PatternFound := FALSE;
IF ExpectedLength = USINT_TO_DINT(Length) THEN
    LastCandidateOffset := 0;
    FOR CandidateOffset := 0 TO LastCandidateOffset DO
        PatternMatches := TRUE;
        FOR CharacterIndex := 0 TO ExpectedLength - 1 DO
            InIndex := LINT_TO_DINT(DINT_TO_LINT(StartIndex) + CandidateOffset
                + DINT_TO_LINT(CharacterIndex));
            IF IN[InIndex] <> Expected[CharacterIndex] THEN
                PatternMatches := FALSE;
                EXIT;
            END_IF;
        END_FOR;
        IF PatternMatches THEN
            PatternFound := TRUE;
            EXIT;
        END_IF;
    END_FOR;
END_IF;

IF NOT PatternFound THEN
    ExpectedText := CreateAssertionTextValue_WString(Value := Expected);
    Message := CONCAT('Assertion failed: selected array does not equal Expected = ',
        ExpectedText);
    Message := CONCAT(Message, ', Range = [');
    Message := CONCAT(Message, DINT_TO_STRING(StartIndex));
    Message := CONCAT(Message, '..');
    Message := CONCAT(Message, LINT_TO_STRING(EndIndex));
    Message := CONCAT(Message, '], ExpectedLength = ');
    Message := CONCAT(Message, DINT_TO_STRING(ExpectedLength));
    Message := CONCAT(Message, '.');
    Fail(Message := Message);
    RETURN;
END_IF;

Pass();
{warning restore C0371}
END_METHOD

END_FUNCTION_BLOCK

// ---- Framework/Assertions/POU/Utilities/IsAssertionWStringLengthValid.TcPOU
{region 'Documentation'}
(*!
<summary>Checks for a terminator within the configured content capacity, including empty text. Reads at most capacity + 1 code units and stops at the first terminator.</summary>
*)
{endregion}
FUNCTION INTERNAL IsAssertionWStringLengthValid : BOOL //! TRUE when a terminator occurs within the configured capacity, including empty text.
VAR_IN_OUT CONSTANT
    Value : WSTRING(Param_Assertions.AssertionWStringLength); //! Read-only text to check for termination within its configured capacity.
END_VAR
VAR
    CharacterIndex : DINT;
END_VAR
VAR CONSTANT
    Terminator : WORD := 0;
END_VAR

IsAssertionWStringLengthValid := FALSE;
FOR CharacterIndex := 0 TO UINT_TO_DINT(Param_Assertions.AssertionWStringLength) DO
    IF Value[CharacterIndex] = Terminator THEN
        IsAssertionWStringLengthValid := TRUE;
        RETURN;
    END_IF;
END_FOR;

END_FUNCTION

// ---- Framework/Assertions/POU/Arrays/Word/AssertArrayContainsWString_Word.TcPOU
{region 'Documentation'}
(*!
<summary>Search the selected array for the contiguous WSTRING code units.</summary>
<description>

StartIndex is an absolute declared IN index, not an offset. Length selects 1..255
elements; the complete selected range must fit IN. Invalid references or ranges report
Error.

Keep supplied arrays stable for the call. Input data is read, not copied or retained as a
snapshot.

Expected must be nonempty and fit its configured text capacity (otherwise Error). A valid
text longer than the selected array region reports Failed. The array is not zero-terminated or
trimmed; matching is exact and case-sensitive.

</description>
*)
{endregion}
FUNCTION_BLOCK AssertArrayContainsWString_Word EXTENDS AssertionBase
VAR_INPUT
    StartIndex : DINT; //! First selected index in IN; uses the array's declared index range, not a zero-based offset.
    Length : USINT; //! Number of selected array elements, from 1 through 255.
END_VAR
VAR_IN_OUT CONSTANT
    IN : ARRAY[*] OF WORD; //! Read-only actual data; the selected range must remain stable during the call.
    Expected : WSTRING(Param_Assertions.AssertionWStringLength); //! Nonempty expected text, terminated within the configured capacity; keep stable during the call.
END_VAR

SUPER^();

{region 'Documentation'}
(*!
<summary>Validate references and ranges before exact code-unit comparison.</summary>
*)
{endregion}
METHOD PROTECTED Assert
VAR
    InLowerIndex : DINT;
    InUpperIndex : DINT;
    EndIndex : LINT;
    ExpectedLength : DINT;
    CharacterIndex : DINT;
    InIndex : DINT;
    CandidateOffset : LINT;
    LastCandidateOffset : LINT;
    PatternMatches : BOOL;
    PatternFound : BOOL;
    ExpectedText : STRING(GVL_Constants.AssertionValueLength);
    Message : STRING(GVL_Constants.MessageLength);
END_VAR
VAR CONSTANT
    Terminator : WORD := 0;
END_VAR
IF NOT EvaluationActive THEN
    RETURN;
END_IF;

IF Result = E_Result.Error THEN
    RETURN;
END_IF;

// C0371: FB inputs are checked before any reference access.
{warning disable C0371}
IF NOT __ISVALIDREF(IN) THEN
    Error(Message := 'Assertion error: IN reference is invalid.');
    RETURN;
END_IF;

IF NOT __ISVALIDREF(Expected) THEN
    Error(Message := 'Assertion error: Expected reference is invalid.');
    RETURN;
END_IF;

IF NOT IsAssertionWStringLengthValid(Value := Expected) THEN
    Error(Message := 'Assertion error: Expected exceeds configured WSTRING length.');
    RETURN;
END_IF;

IF Expected[0] = Terminator THEN
    Error(Message := 'Assertion error: Expected must not be empty.');
    RETURN;
END_IF;

ExpectedLength := 0;
FOR CharacterIndex := 0 TO UINT_TO_DINT(Param_Assertions.AssertionWStringLength) DO
    IF Expected[CharacterIndex] = Terminator THEN
        ExpectedLength := CharacterIndex;
        EXIT;
    END_IF;
END_FOR;

InLowerIndex := LOWER_BOUND(IN, 1);
InUpperIndex := UPPER_BOUND(IN, 1);
EndIndex := DINT_TO_LINT(StartIndex) + USINT_TO_LINT(Length) - 1;
IF (Length = 0)
    OR (StartIndex < InLowerIndex) OR (StartIndex > InUpperIndex)
    OR (EndIndex > DINT_TO_LINT(InUpperIndex)) THEN
    Message := CONCAT('Assertion error: array range is invalid. StartIndex = ',
        DINT_TO_STRING(StartIndex));
    Message := CONCAT(Message, ', Length = ');
    Message := CONCAT(Message, USINT_TO_STRING(Length));
    Error(Message := Message);
    RETURN;
END_IF;

IF Result = E_Result.Failed THEN
    RETURN;
END_IF;

PatternFound := FALSE;
IF ExpectedLength <= USINT_TO_DINT(Length) THEN
    LastCandidateOffset := USINT_TO_LINT(Length) - DINT_TO_LINT(ExpectedLength);
    FOR CandidateOffset := 0 TO LastCandidateOffset DO
        PatternMatches := TRUE;
        FOR CharacterIndex := 0 TO ExpectedLength - 1 DO
            InIndex := LINT_TO_DINT(DINT_TO_LINT(StartIndex) + CandidateOffset
                + DINT_TO_LINT(CharacterIndex));
            IF IN[InIndex] <> Expected[CharacterIndex] THEN
                PatternMatches := FALSE;
                EXIT;
            END_IF;
        END_FOR;
        IF PatternMatches THEN
            PatternFound := TRUE;
            EXIT;
        END_IF;
    END_FOR;
END_IF;

IF NOT PatternFound THEN
    ExpectedText := CreateAssertionTextValue_WString(Value := Expected);
    Message := CONCAT('Assertion failed: selected array does not contain Expected = ',
        ExpectedText);
    Message := CONCAT(Message, ', Range = [');
    Message := CONCAT(Message, DINT_TO_STRING(StartIndex));
    Message := CONCAT(Message, '..');
    Message := CONCAT(Message, LINT_TO_STRING(EndIndex));
    Message := CONCAT(Message, '], ExpectedLength = ');
    Message := CONCAT(Message, DINT_TO_STRING(ExpectedLength));
    Message := CONCAT(Message, '.');
    Fail(Message := Message);
    RETURN;
END_IF;

Pass();
{warning restore C0371}
END_METHOD

END_FUNCTION_BLOCK

// ---- Framework/Assertions/POU/Arrays/Word/AssertArrayStartsWithWString_Word.TcPOU
{region 'Documentation'}
(*!
<summary>Check that the selected array starts with the WSTRING code units.</summary>
<description>

StartIndex is an absolute declared IN index, not an offset. Length selects 1..255
elements; the complete selected range must fit IN. Invalid references or ranges report
Error.

Keep supplied arrays stable for the call. Input data is read, not copied or retained as a
snapshot.

Expected must be nonempty and fit its configured text capacity (otherwise Error). A valid
text longer than the selected array region reports Failed. The array is not zero-terminated or
trimmed; matching is exact and case-sensitive.

</description>
*)
{endregion}
FUNCTION_BLOCK AssertArrayStartsWithWString_Word EXTENDS AssertionBase
VAR_INPUT
    StartIndex : DINT; //! First selected index in IN; uses the array's declared index range, not a zero-based offset.
    Length : USINT; //! Number of selected array elements, from 1 through 255.
END_VAR
VAR_IN_OUT CONSTANT
    IN : ARRAY[*] OF WORD; //! Read-only actual data; the selected range must remain stable during the call.
    Expected : WSTRING(Param_Assertions.AssertionWStringLength); //! Nonempty expected text, terminated within the configured capacity; keep stable during the call.
END_VAR

SUPER^();

{region 'Documentation'}
(*!
<summary>Validate references and ranges before exact code-unit comparison.</summary>
*)
{endregion}
METHOD PROTECTED Assert
VAR
    InLowerIndex : DINT;
    InUpperIndex : DINT;
    EndIndex : LINT;
    ExpectedLength : DINT;
    CharacterIndex : DINT;
    InIndex : DINT;
    CandidateOffset : LINT;
    LastCandidateOffset : LINT;
    PatternMatches : BOOL;
    PatternFound : BOOL;
    ExpectedText : STRING(GVL_Constants.AssertionValueLength);
    Message : STRING(GVL_Constants.MessageLength);
END_VAR
VAR CONSTANT
    Terminator : WORD := 0;
END_VAR
IF NOT EvaluationActive THEN
    RETURN;
END_IF;

IF Result = E_Result.Error THEN
    RETURN;
END_IF;

// C0371: FB inputs are checked before any reference access.
{warning disable C0371}
IF NOT __ISVALIDREF(IN) THEN
    Error(Message := 'Assertion error: IN reference is invalid.');
    RETURN;
END_IF;

IF NOT __ISVALIDREF(Expected) THEN
    Error(Message := 'Assertion error: Expected reference is invalid.');
    RETURN;
END_IF;

IF NOT IsAssertionWStringLengthValid(Value := Expected) THEN
    Error(Message := 'Assertion error: Expected exceeds configured WSTRING length.');
    RETURN;
END_IF;

IF Expected[0] = Terminator THEN
    Error(Message := 'Assertion error: Expected must not be empty.');
    RETURN;
END_IF;

ExpectedLength := 0;
FOR CharacterIndex := 0 TO UINT_TO_DINT(Param_Assertions.AssertionWStringLength) DO
    IF Expected[CharacterIndex] = Terminator THEN
        ExpectedLength := CharacterIndex;
        EXIT;
    END_IF;
END_FOR;

InLowerIndex := LOWER_BOUND(IN, 1);
InUpperIndex := UPPER_BOUND(IN, 1);
EndIndex := DINT_TO_LINT(StartIndex) + USINT_TO_LINT(Length) - 1;
IF (Length = 0)
    OR (StartIndex < InLowerIndex) OR (StartIndex > InUpperIndex)
    OR (EndIndex > DINT_TO_LINT(InUpperIndex)) THEN
    Message := CONCAT('Assertion error: array range is invalid. StartIndex = ',
        DINT_TO_STRING(StartIndex));
    Message := CONCAT(Message, ', Length = ');
    Message := CONCAT(Message, USINT_TO_STRING(Length));
    Error(Message := Message);
    RETURN;
END_IF;

IF Result = E_Result.Failed THEN
    RETURN;
END_IF;

PatternFound := FALSE;
IF ExpectedLength <= USINT_TO_DINT(Length) THEN
    LastCandidateOffset := 0;
    FOR CandidateOffset := 0 TO LastCandidateOffset DO
        PatternMatches := TRUE;
        FOR CharacterIndex := 0 TO ExpectedLength - 1 DO
            InIndex := LINT_TO_DINT(DINT_TO_LINT(StartIndex) + CandidateOffset
                + DINT_TO_LINT(CharacterIndex));
            IF IN[InIndex] <> Expected[CharacterIndex] THEN
                PatternMatches := FALSE;
                EXIT;
            END_IF;
        END_FOR;
        IF PatternMatches THEN
            PatternFound := TRUE;
            EXIT;
        END_IF;
    END_FOR;
END_IF;

IF NOT PatternFound THEN
    ExpectedText := CreateAssertionTextValue_WString(Value := Expected);
    Message := CONCAT('Assertion failed: selected array does not start with Expected = ',
        ExpectedText);
    Message := CONCAT(Message, ', Range = [');
    Message := CONCAT(Message, DINT_TO_STRING(StartIndex));
    Message := CONCAT(Message, '..');
    Message := CONCAT(Message, LINT_TO_STRING(EndIndex));
    Message := CONCAT(Message, '], ExpectedLength = ');
    Message := CONCAT(Message, DINT_TO_STRING(ExpectedLength));
    Message := CONCAT(Message, '.');
    Fail(Message := Message);
    RETURN;
END_IF;

Pass();
{warning restore C0371}
END_METHOD

END_FUNCTION_BLOCK

// ---- Framework/Assertions/POU/Arrays/Word/AssertArrayEndsWithWString_Word.TcPOU
{region 'Documentation'}
(*!
<summary>Check that the selected array ends with the WSTRING code units.</summary>
<description>

StartIndex is an absolute declared IN index, not an offset. Length selects 1..255
elements; the complete selected range must fit IN. Invalid references or ranges report
Error.

Keep supplied arrays stable for the call. Input data is read, not copied or retained as a
snapshot.

Expected must be nonempty and fit its configured text capacity (otherwise Error). A valid
text longer than the selected array region reports Failed. The array is not zero-terminated or
trimmed; matching is exact and case-sensitive.

</description>
*)
{endregion}
FUNCTION_BLOCK AssertArrayEndsWithWString_Word EXTENDS AssertionBase
VAR_INPUT
    StartIndex : DINT; //! First selected index in IN; uses the array's declared index range, not a zero-based offset.
    Length : USINT; //! Number of selected array elements, from 1 through 255.
END_VAR
VAR_IN_OUT CONSTANT
    IN : ARRAY[*] OF WORD; //! Read-only actual data; the selected range must remain stable during the call.
    Expected : WSTRING(Param_Assertions.AssertionWStringLength); //! Nonempty expected text, terminated within the configured capacity; keep stable during the call.
END_VAR

SUPER^();

{region 'Documentation'}
(*!
<summary>Validate references and ranges before exact code-unit comparison.</summary>
*)
{endregion}
METHOD PROTECTED Assert
VAR
    InLowerIndex : DINT;
    InUpperIndex : DINT;
    EndIndex : LINT;
    ExpectedLength : DINT;
    CharacterIndex : DINT;
    InIndex : DINT;
    CandidateOffset : LINT;
    LastCandidateOffset : LINT;
    PatternMatches : BOOL;
    PatternFound : BOOL;
    ExpectedText : STRING(GVL_Constants.AssertionValueLength);
    Message : STRING(GVL_Constants.MessageLength);
END_VAR
VAR CONSTANT
    Terminator : WORD := 0;
END_VAR
IF NOT EvaluationActive THEN
    RETURN;
END_IF;

IF Result = E_Result.Error THEN
    RETURN;
END_IF;

// C0371: FB inputs are checked before any reference access.
{warning disable C0371}
IF NOT __ISVALIDREF(IN) THEN
    Error(Message := 'Assertion error: IN reference is invalid.');
    RETURN;
END_IF;

IF NOT __ISVALIDREF(Expected) THEN
    Error(Message := 'Assertion error: Expected reference is invalid.');
    RETURN;
END_IF;

IF NOT IsAssertionWStringLengthValid(Value := Expected) THEN
    Error(Message := 'Assertion error: Expected exceeds configured WSTRING length.');
    RETURN;
END_IF;

IF Expected[0] = Terminator THEN
    Error(Message := 'Assertion error: Expected must not be empty.');
    RETURN;
END_IF;

ExpectedLength := 0;
FOR CharacterIndex := 0 TO UINT_TO_DINT(Param_Assertions.AssertionWStringLength) DO
    IF Expected[CharacterIndex] = Terminator THEN
        ExpectedLength := CharacterIndex;
        EXIT;
    END_IF;
END_FOR;

InLowerIndex := LOWER_BOUND(IN, 1);
InUpperIndex := UPPER_BOUND(IN, 1);
EndIndex := DINT_TO_LINT(StartIndex) + USINT_TO_LINT(Length) - 1;
IF (Length = 0)
    OR (StartIndex < InLowerIndex) OR (StartIndex > InUpperIndex)
    OR (EndIndex > DINT_TO_LINT(InUpperIndex)) THEN
    Message := CONCAT('Assertion error: array range is invalid. StartIndex = ',
        DINT_TO_STRING(StartIndex));
    Message := CONCAT(Message, ', Length = ');
    Message := CONCAT(Message, USINT_TO_STRING(Length));
    Error(Message := Message);
    RETURN;
END_IF;

IF Result = E_Result.Failed THEN
    RETURN;
END_IF;

PatternFound := FALSE;
IF ExpectedLength <= USINT_TO_DINT(Length) THEN
    LastCandidateOffset := USINT_TO_LINT(Length) - DINT_TO_LINT(ExpectedLength);
    FOR CandidateOffset := USINT_TO_LINT(Length) - DINT_TO_LINT(ExpectedLength) TO LastCandidateOffset DO
        PatternMatches := TRUE;
        FOR CharacterIndex := 0 TO ExpectedLength - 1 DO
            InIndex := LINT_TO_DINT(DINT_TO_LINT(StartIndex) + CandidateOffset
                + DINT_TO_LINT(CharacterIndex));
            IF IN[InIndex] <> Expected[CharacterIndex] THEN
                PatternMatches := FALSE;
                EXIT;
            END_IF;
        END_FOR;
        IF PatternMatches THEN
            PatternFound := TRUE;
            EXIT;
        END_IF;
    END_FOR;
END_IF;

IF NOT PatternFound THEN
    ExpectedText := CreateAssertionTextValue_WString(Value := Expected);
    Message := CONCAT('Assertion failed: selected array does not end with Expected = ',
        ExpectedText);
    Message := CONCAT(Message, ', Range = [');
    Message := CONCAT(Message, DINT_TO_STRING(StartIndex));
    Message := CONCAT(Message, '..');
    Message := CONCAT(Message, LINT_TO_STRING(EndIndex));
    Message := CONCAT(Message, '], ExpectedLength = ');
    Message := CONCAT(Message, DINT_TO_STRING(ExpectedLength));
    Message := CONCAT(Message, '.');
    Fail(Message := Message);
    RETURN;
END_IF;

Pass();
{warning restore C0371}
END_METHOD

END_FUNCTION_BLOCK

// ---- SelfTests/TestSuites/TestSuite_AssertionVariants.TcPOU
{region 'Documentation'}
(*!
<summary>Checks selected residual Assertion operators, operand widths and diagnostics.</summary>
*)
{endregion}
FUNCTION_BLOCK TestSuite_AssertionVariants EXTENDS TestSuiteBase
VAR
    FBitSelection : Test_AssertionBitSelection;
    FMaskPredicates : Test_AssertionMaskPredicates;
    FCountPredicates : Test_AssertionCountPredicates;
    FNarrowIntegers : Test_AssertionNarrowIntegers;
    FTemporalVariants : Test_AssertionTemporalVariants;
    FTestCases : ARRAY[1..TestCaseCapacity] OF I_TestCase;
END_VAR
VAR CONSTANT
    TestCaseCapacity : UINT := 5;
END_VAR

SUPER^();

{region 'Documentation'}
(*!
<summary>Initializes five focused residual Assertion Test Cases and registers them serially.</summary>
*)
{endregion}
METHOD PROTECTED Configure
VAR_IN_OUT
    // SA0167: Borrowed owner builder; no temporary instance is created.
    {attribute 'analysis' := '-167'}
    Builder : TestSuiteConfigurationBuilder; //! Borrowed owner configuration builder used only during this Configure call; register this owner's concrete children.
END_VAR
VAR
    TestConfig : ST_TestCaseConfig;
END_VAR
Builder.Initialize(Mode := E_OrchestrationMode.Serial,
    TestCases := FTestCases);
FBitSelection.Initialize(Parent := THIS^,
    TestName := 'BitSelection',
    Config := TestConfig);
Builder.Register(TestCase := FBitSelection);
FMaskPredicates.Initialize(Parent := THIS^,
    TestName := 'MaskPredicates',
    Config := TestConfig);
Builder.Register(TestCase := FMaskPredicates);
FCountPredicates.Initialize(Parent := THIS^,
    TestName := 'CountPredicates',
    Config := TestConfig);
Builder.Register(TestCase := FCountPredicates);
FNarrowIntegers.Initialize(Parent := THIS^,
    TestName := 'NarrowIntegers',
    Config := TestConfig);
Builder.Register(TestCase := FNarrowIntegers);
FTemporalVariants.Initialize(Parent := THIS^,
    TestName := 'TemporalVariants',
    Config := TestConfig);
Builder.Register(TestCase := FTemporalVariants);
END_METHOD

{region 'Documentation'}
(*!
<summary>Returns a registered scenario using its original array index.</summary>
*)
{endregion}
METHOD PUBLIC GetTestCase : I_TestCase //! Typed child interface at the original array index; zero when no entry is available.
VAR_INPUT
    Index : DINT; //! Original occupied child-array index, rather than an ordinal position.
END_VAR
GetTestCase := 0;
IF (ChildCount = 0) OR (Index < ChildArrayLowerBound)
    OR (DINT_TO_LINT(Index) >= DINT_TO_LINT(ChildArrayLowerBound) + UINT_TO_LINT(ChildCount)) THEN
    RETURN;
END_IF;
GetTestCase := FTestCases[Index];
END_METHOD

{region 'Documentation'}
(*!
<summary>Calls every owned scenario once per initialized Suite cycle.</summary>
*)
{endregion}
METHOD PROTECTED ProcessTestCases
FBitSelection();
FMaskPredicates();
FCountPredicates();
FNarrowIntegers();
FTemporalVariants();
END_METHOD

END_FUNCTION_BLOCK

// ---- SelfTests/TestCases/TestSuite_AssertionVariants/Test_AssertionBitSelection.TcPOU
{region 'Documentation'}
(*!
<summary>Checks bit selection with isolated production subjects.</summary>
<description>
Each independent scenario consumes a bound reset call before its evaluation call.
ProcessAssertions checks the observation before ProcessTests advances.
SelectScenario holds explicit expected results; no production algorithm is mirrored.
Expected findings remain in the local capture; only outer checks affect the test result.
FirstFailedScenario and FailedDuringEvaluation retain the first mismatch.
The final scenario retains Failed and changes only the bit indices on the next call; Error must still escalate.
</description>
*)
{endregion}
FUNCTION_BLOCK Test_AssertionBitSelection EXTENDS TestCaseBase
VAR
    FTrueBit : AssertTrueBit_LWord;
    FTrueBitExpectedResult : E_Result;
    FTrueBitExpectedFinding : BOOL;
    FNotEqualBit : AssertNotEqualBit_Byte;
    FNotEqualBitExpectedResult : E_Result;
    FNotEqualBitExpectedFinding : BOOL;

    FWideValue : LWORD;
    FByteValue : BYTE;
    FWideIndex : USINT;
    FByteIndex : USINT;
    FForbidden : BOOL;
    FEscalating : BOOL;
    FSubjectEnable : BOOL;
    FCapture : EventBuffer;
    FEvents : ARRAY[1..CaptureLength] OF ST_Event;
    FCaptureFifo : ST_FifoStatus;
    FCaptureStatus : ST_EventBufferStatus;
    FSetupValid : BOOL;
    FScenario : UINT;
    FChecked : BOOL;
    FEvaluateSubjects : BOOL;
    FObservationReady : BOOL;
    FFirstFailedScenario : UINT;
    FFailedDuringEvaluation : BOOL;
    FResultsMatch : BOOL;
    FResults : AssertTrue;
    FActivityMatch : BOOL;
    FActivity : AssertTrue;
    FInputsMatch : BOOL;
    FInputs : AssertTrue;
    FFindingsMatch : BOOL;
    FFindings : AssertTrue;
END_VAR
VAR CONSTANT
    CaptureLength : UINT := 8;
    ScenarioLowestBit : UINT := 1;
    ScenarioHighestBit : UINT := 2;
    ScenarioAdjacentBit : UINT := 3;
    ScenarioForbiddenTrue : UINT := 4;
    ScenarioInvalidIndex : UINT := 5;
    ScenarioFailedThenError : UINT := 6;
    LastScenario : UINT := ScenarioFailedThenError;
END_VAR

SUPER^();

{region 'Documentation'}
(*!
<summary>Aggregates only outer checks, not intentionally failing subjects.</summary>
*)
{endregion}
METHOD PROTECTED AggregateResults
VAR_INPUT
    Aggregator : I_ResultAggregator; //! Borrowed result sink owned by the outer Test Case; add this test's checking Assertions without resetting or retaining the sink.
END_VAR
Aggregator.AddProvider(Provider := FResults);
Aggregator.AddProvider(Provider := FActivity);
Aggregator.AddProvider(Provider := FInputs);
Aggregator.AddProvider(Provider := FFindings);
END_METHOD

{region 'Documentation'}
(*!
<summary>Calls each inherited production subject once with caller-owned input storage.</summary>
*)
{endregion}
METHOD PRIVATE CallSubjects
FTrueBit(Enable := FSubjectEnable,
    State := E_State.Running,
    IN := FWideValue,
    BitIndex := FWideIndex);
FNotEqualBit(Enable := FSubjectEnable,
    State := E_State.Running,
    IN := FByteValue,
    BitIndex := FByteIndex,
    Expected := FForbidden);
END_METHOD

{region 'Documentation'}
(*!
<summary>Checks one subject finding in call order; expected outcomes come from the scenario.</summary>
*)
{endregion}
METHOD PRIVATE CheckFinding : BOOL //! TRUE when the required finding checks pass; calls requiring no finding also succeed.
VAR_INPUT
    Subject : I_Assertion; //! Assertion interface supplying the expected finding identity.
    ExpectedResult : E_Result; //! Independently authored result expected in the captured finding.
    ExpectedFinding : BOOL; //! TRUE when this scenario requires a finding during active evaluation.
END_VAR
VAR_IN_OUT
    Index : UINT; //! One-based next finding index; advanced when this call checks a required finding.
END_VAR
CheckFinding := TRUE;
IF FEvaluateSubjects AND ExpectedFinding THEN
    CheckFinding := (FEvents[Index].SequenceId = UINT_TO_UDINT(Index))
        AND (FEvents[Index].Name = Subject.Name)
        AND (FEvents[Index].OwnerScope = E_OwnerScope.Assertion)
        AND (FEvents[Index].EventType = E_EventType.Result)
        AND (FEvents[Index].State = E_State.Running)
        AND (FEvents[Index].Result = ExpectedResult)
        AND (FEvents[Index].Message <> '');
    Index := Index + 1;
END_IF;
END_METHOD

{region 'Documentation'}
(*!
<summary>Checks exact finding count and identities; at most one finding per subject.</summary>
*)
{endregion}
METHOD PRIVATE CheckFindings
VAR
    Index : UINT;
    Matches : BOOL;
END_VAR
Index := 1;
FFindingsMatch := TRUE;
Matches := CheckFinding(Subject := FTrueBit,
    ExpectedResult := FTrueBitExpectedResult,
    ExpectedFinding := FTrueBitExpectedFinding,
    Index := Index);
FFindingsMatch := FFindingsMatch AND Matches;
Matches := CheckFinding(Subject := FNotEqualBit,
    ExpectedResult := FNotEqualBitExpectedResult,
    ExpectedFinding := FNotEqualBitExpectedFinding,
    Index := Index);
FFindingsMatch := FFindingsMatch AND Matches;
FFindingsMatch := FFindingsMatch
    AND (FCaptureStatus.SequenceId = UINT_TO_UDINT(Index - 1))
    AND (FCaptureStatus.LostEventCount = 0);
IF FEvaluateSubjects AND (FScenario = ScenarioAdjacentBit) THEN
    // SA0175: Fixed byte-substring checks of bounded diagnostic messages; no character offsets.
    {analysis -175}
    FFindingsMatch := FFindingsMatch
        AND (FIND(FEvents[1].Message, 'BitIndex = 63') > 0)
        AND (FIND(FEvents[2].Message, 'BitIndex = 7') > 0)
        AND (FIND(FEvents[2].Message, 'Value = 16#40') > 0);
    {analysis +175}
END_IF;
END_METHOD

{region 'Documentation'}
(*!
<summary>Rejects incomplete subject, capture or outer Assertion setup.</summary>
*)
{endregion}
METHOD PROTECTED CheckInitialization : BOOL //! TRUE when the inherited initialization check and this concrete fixture check both accept the setup.
CheckInitialization := SUPER^.CheckInitialization();
IF NOT CheckInitialization THEN
    RETURN;
END_IF;

CheckInitialization := FSetupValid
    AND FResults.IsInitialized
    AND FActivity.IsInitialized
    AND FInputs.IsInitialized
    AND FFindings.IsInitialized;
IF NOT CheckInitialization THEN
    EventPublisher.PublishEvent(Event := CreateFrameworkEvent(Name := Name,
        ResourceName := '',
        State := State,
        Severity := E_EventSeverity.Error,
        Message := 'Variant selftest setup failed.'));
END_IF;
END_METHOD

{region 'Documentation'}
(*!
<summary>Verifies input preservation without using the tested comparison algorithm.</summary>
*)
{endregion}
METHOD PRIVATE CheckInputs
FInputsMatch := (FTrueBit.IN = FWideValue)
    AND (FTrueBit.BitIndex = FWideIndex)
    AND (FNotEqualBit.IN = FByteValue)
    AND (FNotEqualBit.BitIndex = FByteIndex)
    AND (FNotEqualBit.Expected = FForbidden);
END_METHOD

{region 'Documentation'}
(*!
<summary>Checks literal evaluation results, or NotEvaluated on the reset call.</summary>
*)
{endregion}
METHOD PRIVATE CheckResults
IF FEvaluateSubjects THEN
    FResultsMatch := (FTrueBit.Result = FTrueBitExpectedResult)
        AND (FNotEqualBit.Result = FNotEqualBitExpectedResult);
ELSE
    FResultsMatch := (FTrueBit.Result = E_Result.NotEvaluated)
        AND (FNotEqualBit.Result = E_Result.NotEvaluated);
END_IF;
FActivityMatch := (FTrueBit.Enabled = FSubjectEnable)
    AND (FTrueBit.ObservationActive = (FEvaluateSubjects AND FSubjectEnable))
    AND (FTrueBit.EvaluationActive = (FEvaluateSubjects AND FSubjectEnable))
    AND (FNotEqualBit.Enabled = FSubjectEnable)
    AND (FNotEqualBit.ObservationActive = (FEvaluateSubjects AND FSubjectEnable))
    AND (FNotEqualBit.EvaluationActive = (FEvaluateSubjects AND FSubjectEnable));
END_METHOD

{region 'Documentation'}
(*!
<summary>Initializes outer checks and isolates intentional subject findings.</summary>
*)
{endregion}
METHOD PROTECTED Configure
VAR
    Initialized : BOOL;
END_VAR
FPreparationStateCount := 0;
FTestStateCount := 1;
FResults.Initialize(Parent := THIS^,
    AssertionName := 'Results');
FActivity.Initialize(Parent := THIS^,
    AssertionName := 'Activity');
FInputs.Initialize(Parent := THIS^,
    AssertionName := 'Inputs');
FFindings.Initialize(Parent := THIS^,
    AssertionName := 'Findings');
FSetupValid := FCapture.Initialize(Buffer := FEvents,
    FifoControl := FCaptureFifo,
    Status := FCaptureStatus);
FTrueBit.BindPublisher(Publisher := FCapture);
Initialized := FTrueBit.Initialize(Parent := THIS^,
    AssertionName := 'TrueBit');
FSetupValid := FSetupValid AND Initialized;
FNotEqualBit.BindPublisher(Publisher := FCapture);
Initialized := FNotEqualBit.Initialize(Parent := THIS^,
    AssertionName := 'NotEqualBit');
FSetupValid := FSetupValid AND Initialized;
END_METHOD

{region 'Documentation'}
(*!
<summary>Completes abort; no asynchronous resource is owned.</summary>
*)
{endregion}
METHOD PROTECTED ProcessAbort
VAR_INPUT
    Enable : BOOL; //! Phase permission supplied by the owning Test Case; FALSE does not authorize progression, while observation may continue.
END_VAR
IF Enable THEN
    CompleteAbort();
END_IF;
END_METHOD

{region 'Documentation'}
(*!
<summary>Latches this call's checks before progression is permitted.</summary>
*)
{endregion}
METHOD PROTECTED ProcessAssertions
VAR_INPUT
    Enable : BOOL; //! Phase permission supplied by the owning Test Case; FALSE does not authorize progression, while observation may continue.
END_VAR
VAR
    Check : BOOL;
END_VAR
Check := Enable AND FObservationReady;
FResults(Enable := Check,
    State := State,
    IN := FResultsMatch);
FActivity(Enable := Check,
    State := State,
    IN := FActivityMatch);
FInputs(Enable := Check,
    State := State,
    IN := FInputsMatch);
FFindings(Enable := Check,
    State := State,
    IN := FFindingsMatch);
IF Check THEN
    FChecked := TRUE;
END_IF;
END_METHOD

{region 'Documentation'}
(*!
<summary>No Preparation phase is needed.</summary>
*)
{endregion}
METHOD PROTECTED ProcessPreparations
VAR_INPUT
    // SA0033: Required hook; this test has no Preparation phase.
    {attribute 'analysis' := '-33'}
    Enable : BOOL; //! Phase permission supplied by the owning Test Case; FALSE does not authorize progression, while observation may continue.
END_VAR
END_METHOD

{region 'Documentation'}
(*!
<summary>Restarts the scenario sequence and outer checks.</summary>
*)
{endregion}
METHOD PROTECTED ProcessReset
FScenario := ScenarioLowestBit;
FEscalating := FALSE;
FChecked := FALSE;
FSubjectEnable := FALSE;
FEvaluateSubjects := FALSE;
FObservationReady := FALSE;
FFirstFailedScenario := 0;
FFailedDuringEvaluation := FALSE;
FCapture.Reset();
ResetSubjects();
FResults.Reset();
FActivity.Reset();
FInputs.Reset();
FFindings.Reset();
CompleteReset();
END_METHOD

{region 'Documentation'}
(*!
<summary>Consumes reset, evaluates, then waits for the outer checks before advancing.</summary>
*)
{endregion}
METHOD PROTECTED ProcessTests
VAR_INPUT
    Enable : BOOL; //! Phase permission supplied by the owning Test Case; FALSE does not authorize progression, while observation may continue.
END_VAR
IF NOT Enable THEN
    RETURN;
END_IF;

IF FChecked THEN
    FChecked := FALSE;
    FObservationReady := FALSE;
    IF FEvaluateSubjects THEN
        IF FScenario = LastScenario THEN
            IF FEscalating THEN
                CompleteTests();
                RETURN;
            END_IF;
            FEscalating := TRUE;
        ELSE
            FScenario := FScenario + 1;
        END_IF;
    END_IF;
    FEvaluateSubjects := FEscalating OR NOT FEvaluateSubjects;
END_IF;

IF NOT SelectScenario() THEN
    RETURN;
END_IF;
FCapture.Reset();
IF NOT FEvaluateSubjects THEN
    ResetSubjects();
END_IF;

CallSubjects();
CheckResults();
CheckInputs();
CheckFindings();
IF (FFirstFailedScenario = 0)
    AND NOT (FResultsMatch AND FActivityMatch AND FInputsMatch AND FFindingsMatch) THEN
    FFirstFailedScenario := FScenario;
    FFailedDuringEvaluation := FEvaluateSubjects;
END_IF;
FObservationReady := TRUE;
END_METHOD

{region 'Documentation'}
(*!
<summary>Queues reset; the next bound FB call consumes it without evaluating.</summary>
*)
{endregion}
METHOD PRIVATE ResetSubjects
FTrueBit.Reset();
FNotEqualBit.Reset();
END_METHOD

{region 'Documentation'}
(*!
<summary>Selects explicit stimuli and expected results for one scenario.</summary>
*)
{endregion}
METHOD PRIVATE SelectScenario : BOOL //! TRUE after selecting a supported scenario and its literal expectations; FALSE reports an unknown scenario.
SelectScenario := FALSE;
FSubjectEnable := TRUE;
FWideValue := LWORD#16#0000000000000001;
FByteValue := BYTE#16#01;
FWideIndex := 0;
FByteIndex := 0;
FForbidden := FALSE;
CASE FScenario OF
    ScenarioLowestBit:
        FTrueBitExpectedResult := E_Result.Passed;
        FTrueBitExpectedFinding := FALSE;
        FNotEqualBitExpectedResult := E_Result.Passed;
        FNotEqualBitExpectedFinding := FALSE;
    ScenarioHighestBit:
        FWideValue := LWORD#16#8000000000000000;
        FByteValue := BYTE#16#80;
        FWideIndex := 63;
        FByteIndex := 7;
        FTrueBitExpectedResult := E_Result.Passed;
        FTrueBitExpectedFinding := FALSE;
        FNotEqualBitExpectedResult := E_Result.Passed;
        FNotEqualBitExpectedFinding := FALSE;
    ScenarioAdjacentBit:
        FWideValue := LWORD#16#4000000000000000;
        FByteValue := BYTE#16#40;
        FWideIndex := 63;
        FByteIndex := 7;
        FTrueBitExpectedResult := E_Result.Failed;
        FTrueBitExpectedFinding := TRUE;
        FNotEqualBitExpectedResult := E_Result.Failed;
        FNotEqualBitExpectedFinding := TRUE;
    ScenarioForbiddenTrue:
        FByteValue := 0;
        FForbidden := TRUE;
        FTrueBitExpectedResult := E_Result.Passed;
        FTrueBitExpectedFinding := FALSE;
        FNotEqualBitExpectedResult := E_Result.Passed;
        FNotEqualBitExpectedFinding := FALSE;
    ScenarioInvalidIndex:
        FWideIndex := 64;
        FByteIndex := 8;
        FTrueBitExpectedResult := E_Result.Error;
        FTrueBitExpectedFinding := TRUE;
        FNotEqualBitExpectedResult := E_Result.Error;
        FNotEqualBitExpectedFinding := TRUE;
    ScenarioFailedThenError:
        FWideValue := 0;
        FByteValue := 0;
        FTrueBitExpectedResult := E_Result.Failed;
        FTrueBitExpectedFinding := TRUE;
        FNotEqualBitExpectedResult := E_Result.Failed;
        FNotEqualBitExpectedFinding := TRUE;
ELSE
    Error(Message := 'Unknown variant Assertion scenario.');
    RETURN;
END_CASE;

IF FEscalating THEN
    FWideIndex := 64;
    FByteIndex := 8;
    FTrueBitExpectedResult := E_Result.Error;
    FNotEqualBitExpectedResult := E_Result.Error;
END_IF;
SelectScenario := TRUE;
END_METHOD

END_FUNCTION_BLOCK

// ---- Framework/Assertions/POU/BasicTypes/Byte/AssertNotEqualBit_Byte.TcPOU
{region 'Documentation'}
(*!
<summary>Checks that the selected BYTE bit differs from the expected Boolean value.</summary>
*)
{endregion}
FUNCTION_BLOCK AssertNotEqualBit_Byte EXTENDS AssertionBase
VAR_INPUT
    IN : BYTE; //! Actual bitfield.
    BitIndex : USINT; //! Zero-based bit index (0..7); an invalid index produces Error during evaluation.
    Expected : BOOL; //! Forbidden selected bit value.
END_VAR

SUPER^();

{region 'Documentation'}
(*!
<summary>Validates the index before evaluating the selected bit.</summary>
*)
{endregion}
METHOD PROTECTED Assert
VAR
    Mask : BYTE;
    ActualBit : BOOL;
    Message : STRING(GVL_Constants.MessageLength);
    ActualText : STRING(GVL_Constants.AssertionValueLength);
END_VAR
VAR CONSTANT
    MaxBitIndex : USINT := 7;
    SingleBitMask : BYTE := 16#01;
    NoBitMask : BYTE := 16#00;
    HexDigitCount : USINT := 2;
END_VAR
IF NOT EvaluationActive THEN
    RETURN;
END_IF;

IF Result = E_Result.Error THEN
    RETURN;
END_IF;

IF BitIndex > MaxBitIndex THEN
    Message := CONCAT('Assertion error: bit index is outside valid range. BitIndex = ',
        USINT_TO_STRING(BitIndex));
    Message := CONCAT(Message, ', MaxBitIndex = ');
    Message := CONCAT(Message, USINT_TO_STRING(MaxBitIndex));
    Message := CONCAT(Message, '.');
    Error(Message := Message);
    RETURN;
END_IF;

IF Result = E_Result.Failed THEN
    RETURN;
END_IF;

Mask := SHL(SingleBitMask, BitIndex);
ActualBit := (IN AND Mask) <> NoBitMask;

IF ActualBit = Expected THEN
    ActualText := CreateAssertionTextValue_Hex(Value := BYTE_TO_LWORD(IN),
        DigitCount := HexDigitCount);
    Message := CONCAT('Assertion failed: bit value matches forbidden value. BitIndex = ',
        USINT_TO_STRING(BitIndex));
    Message := CONCAT(Message, ', NotExpected = ');
    Message := CONCAT(Message, BOOL_TO_STRING(Expected));
    Message := CONCAT(Message, ', Actual = ');
    Message := CONCAT(Message, BOOL_TO_STRING(ActualBit));
    Message := CONCAT(Message, ', Value = ');
    Message := CONCAT(Message, ActualText);
    Message := CONCAT(Message, '.');
    Fail(Message := Message);
    RETURN;
END_IF;

Pass();
END_METHOD

END_FUNCTION_BLOCK

// ---- SelfTests/TestCases/TestSuite_AssertionVariants/Test_AssertionMaskPredicates.TcPOU
{region 'Documentation'}
(*!
<summary>Distinguishes masked equality, all-bits and any-bit predicates across bit widths.</summary>
<description>
Each independent scenario consumes a bound reset call before its evaluation call.
ProcessAssertions checks the observation before ProcessTests advances.
SelectScenario holds explicit expected results; no production algorithm is mirrored.
Expected findings remain in the local capture; only outer checks affect the test result.
FirstFailedScenario and FailedDuringEvaluation retain the first mismatch.
Each scenario uses literal typed inputs at the declared operand widths.
</description>
*)
{endregion}
FUNCTION_BLOCK Test_AssertionMaskPredicates EXTENDS TestCaseBase
VAR
    FEqual : AssertEqualMask_Word;
    FEqualExpectedResult : E_Result;
    FEqualExpectedFinding : BOOL;
    FNotEqual : AssertNotEqualMask_LWord;
    FNotEqualExpectedResult : E_Result;
    FNotEqualExpectedFinding : BOOL;
    FAllTrue : AssertTrueMask_Byte;
    FAllTrueExpectedResult : E_Result;
    FAllTrueExpectedFinding : BOOL;
    FAllFalse : AssertFalseMask_DWord;
    FAllFalseExpectedResult : E_Result;
    FAllFalseExpectedFinding : BOOL;
    FContains : AssertContainsBit_LWord;
    FContainsExpectedResult : E_Result;
    FContainsExpectedFinding : BOOL;

    FWordValue : WORD;
    FWordMask : WORD;
    FExpectedWord : WORD;
    FWideValue : LWORD;
    FWideMask : LWORD;
    FForbiddenWide : LWORD;
    FByteValue : BYTE;
    FByteMask : BYTE;
    FDWordValue : DWORD;
    FDWordMask : DWORD;
    FContainsValue : LWORD;
    FContainsMask : LWORD;
    FExpectedBit : BOOL;
    FSubjectEnable : BOOL;
    FCapture : EventBuffer;
    FEvents : ARRAY[1..CaptureLength] OF ST_Event;
    FCaptureFifo : ST_FifoStatus;
    FCaptureStatus : ST_EventBufferStatus;
    FSetupValid : BOOL;
    FScenario : UINT;
    FChecked : BOOL;
    FEvaluateSubjects : BOOL;
    FObservationReady : BOOL;
    FFirstFailedScenario : UINT;
    FFailedDuringEvaluation : BOOL;
    FResultsMatch : BOOL;
    FResults : AssertTrue;
    FActivityMatch : BOOL;
    FActivity : AssertTrue;
    FInputsMatch : BOOL;
    FInputs : AssertTrue;
    FFindingsMatch : BOOL;
    FFindings : AssertTrue;
END_VAR
VAR CONSTANT
    CaptureLength : UINT := 12;
    ScenarioOutsideBitsIgnored : UINT := 1;
    ScenarioPartialSelection : UINT := 2;
    ScenarioContainsFalse : UINT := 3;
    ScenarioAllSelectedTrue : UINT := 4;
    ScenarioAllSelectedFalse : UINT := 5;
    ScenarioFalsePresent : UINT := 6;
    ScenarioEmptyMasks : UINT := 7;
    LastScenario : UINT := ScenarioEmptyMasks;
END_VAR

SUPER^();

{region 'Documentation'}
(*!
<summary>Aggregates only outer checks, not intentionally failing subjects.</summary>
*)
{endregion}
METHOD PROTECTED AggregateResults
VAR_INPUT
    Aggregator : I_ResultAggregator; //! Borrowed result sink owned by the outer Test Case; add this test's checking Assertions without resetting or retaining the sink.
END_VAR
Aggregator.AddProvider(Provider := FResults);
Aggregator.AddProvider(Provider := FActivity);
Aggregator.AddProvider(Provider := FInputs);
Aggregator.AddProvider(Provider := FFindings);
END_METHOD

{region 'Documentation'}
(*!
<summary>Calls each inherited production subject once with caller-owned input storage.</summary>
*)
{endregion}
METHOD PRIVATE CallSubjects
FEqual(Enable := FSubjectEnable,
    State := E_State.Running,
    IN := FWordValue,
    Mask := FWordMask,
    Expected := FExpectedWord);
FNotEqual(Enable := FSubjectEnable,
    State := E_State.Running,
    IN := FWideValue,
    Mask := FWideMask,
    Expected := FForbiddenWide);
FAllTrue(Enable := FSubjectEnable,
    State := E_State.Running,
    IN := FByteValue,
    Mask := FByteMask);
FAllFalse(Enable := FSubjectEnable,
    State := E_State.Running,
    IN := FDWordValue,
    Mask := FDWordMask);
FContains(Enable := FSubjectEnable,
    State := E_State.Running,
    IN := FContainsValue,
    Mask := FContainsMask,
    Expected := FExpectedBit);
END_METHOD

{region 'Documentation'}
(*!
<summary>Checks one subject finding in call order; expected outcomes come from the scenario.</summary>
*)
{endregion}
METHOD PRIVATE CheckFinding : BOOL //! TRUE when the required finding checks pass; calls requiring no finding also succeed.
VAR_INPUT
    Subject : I_Assertion; //! Assertion interface supplying the expected finding identity.
    ExpectedResult : E_Result; //! Independently authored result expected in the captured finding.
    ExpectedFinding : BOOL; //! TRUE when this scenario requires a finding during active evaluation.
END_VAR
VAR_IN_OUT
    Index : UINT; //! One-based next finding index; advanced when this call checks a required finding.
END_VAR
CheckFinding := TRUE;
IF FEvaluateSubjects AND ExpectedFinding THEN
    CheckFinding := (FEvents[Index].SequenceId = UINT_TO_UDINT(Index))
        AND (FEvents[Index].Name = Subject.Name)
        AND (FEvents[Index].OwnerScope = E_OwnerScope.Assertion)
        AND (FEvents[Index].EventType = E_EventType.Result)
        AND (FEvents[Index].State = E_State.Running)
        AND (FEvents[Index].Result = ExpectedResult)
        AND (FEvents[Index].Message <> '');
    Index := Index + 1;
END_IF;
END_METHOD

{region 'Documentation'}
(*!
<summary>Checks exact finding count and identities; at most one finding per subject.</summary>
*)
{endregion}
METHOD PRIVATE CheckFindings
VAR
    Index : UINT;
    Matches : BOOL;
END_VAR
Index := 1;
FFindingsMatch := TRUE;
Matches := CheckFinding(Subject := FEqual,
    ExpectedResult := FEqualExpectedResult,
    ExpectedFinding := FEqualExpectedFinding,
    Index := Index);
FFindingsMatch := FFindingsMatch AND Matches;
Matches := CheckFinding(Subject := FNotEqual,
    ExpectedResult := FNotEqualExpectedResult,
    ExpectedFinding := FNotEqualExpectedFinding,
    Index := Index);
FFindingsMatch := FFindingsMatch AND Matches;
Matches := CheckFinding(Subject := FAllTrue,
    ExpectedResult := FAllTrueExpectedResult,
    ExpectedFinding := FAllTrueExpectedFinding,
    Index := Index);
FFindingsMatch := FFindingsMatch AND Matches;
Matches := CheckFinding(Subject := FAllFalse,
    ExpectedResult := FAllFalseExpectedResult,
    ExpectedFinding := FAllFalseExpectedFinding,
    Index := Index);
FFindingsMatch := FFindingsMatch AND Matches;
Matches := CheckFinding(Subject := FContains,
    ExpectedResult := FContainsExpectedResult,
    ExpectedFinding := FContainsExpectedFinding,
    Index := Index);
FFindingsMatch := FFindingsMatch AND Matches;
FFindingsMatch := FFindingsMatch
    AND (FCaptureStatus.SequenceId = UINT_TO_UDINT(Index - 1))
    AND (FCaptureStatus.LostEventCount = 0);
IF FEvaluateSubjects AND (FScenario = ScenarioPartialSelection) THEN
    // SA0175: Fixed byte-substring checks of bounded diagnostic messages; no character offsets.
    {analysis -175}
    FFindingsMatch := FFindingsMatch
        AND (FIND(FEvents[1].Message, 'Expected = 16#0005') > 0)
        AND (FIND(FEvents[1].Message, 'Mask = 16#00FF') > 0)
        AND (FIND(FEvents[1].Message, 'Actual = 16#A504') > 0)
        AND (FIND(FEvents[2].Message, 'NotExpected = 16#0000000000000000') > 0)
        AND (FIND(FEvents[2].Message, 'Actual = 16#0000000000000001') > 0)
        AND (FIND(FEvents[3].Message, 'Mask = 16#03') > 0)
        AND (FIND(FEvents[3].Message, 'Actual = 16#F1') > 0)
        AND (FIND(FEvents[4].Message, 'Mask = 16#00000003') > 0)
        AND (FIND(FEvents[4].Message, 'Actual = 16#80000001') > 0);
    {analysis +175}
END_IF;
END_METHOD

{region 'Documentation'}
(*!
<summary>Rejects incomplete subject, capture or outer Assertion setup.</summary>
*)
{endregion}
METHOD PROTECTED CheckInitialization : BOOL //! TRUE when the inherited initialization check and this concrete fixture check both accept the setup.
CheckInitialization := SUPER^.CheckInitialization();
IF NOT CheckInitialization THEN
    RETURN;
END_IF;

CheckInitialization := FSetupValid
    AND FResults.IsInitialized
    AND FActivity.IsInitialized
    AND FInputs.IsInitialized
    AND FFindings.IsInitialized;
IF NOT CheckInitialization THEN
    EventPublisher.PublishEvent(Event := CreateFrameworkEvent(Name := Name,
        ResourceName := '',
        State := State,
        Severity := E_EventSeverity.Error,
        Message := 'Variant selftest setup failed.'));
END_IF;
END_METHOD

{region 'Documentation'}
(*!
<summary>Verifies input preservation without using the tested comparison algorithm.</summary>
*)
{endregion}
METHOD PRIVATE CheckInputs
FInputsMatch := (FEqual.IN = FWordValue)
    AND (FEqual.Mask = FWordMask) AND (FEqual.Expected = FExpectedWord)
    AND (FNotEqual.IN = FWideValue)
    AND (FNotEqual.Mask = FWideMask) AND (FNotEqual.Expected = FForbiddenWide)
    AND (FAllTrue.IN = FByteValue) AND (FAllTrue.Mask = FByteMask)
    AND (FAllFalse.IN = FDWordValue) AND (FAllFalse.Mask = FDWordMask)
    AND (FContains.IN = FContainsValue)
    AND (FContains.Mask = FContainsMask) AND (FContains.Expected = FExpectedBit);
END_METHOD

{region 'Documentation'}
(*!
<summary>Checks literal evaluation results, or NotEvaluated on the reset call.</summary>
*)
{endregion}
METHOD PRIVATE CheckResults
IF FEvaluateSubjects THEN
    FResultsMatch := (FEqual.Result = FEqualExpectedResult)
        AND (FNotEqual.Result = FNotEqualExpectedResult)
        AND (FAllTrue.Result = FAllTrueExpectedResult)
        AND (FAllFalse.Result = FAllFalseExpectedResult)
        AND (FContains.Result = FContainsExpectedResult);
ELSE
    FResultsMatch := (FEqual.Result = E_Result.NotEvaluated)
        AND (FNotEqual.Result = E_Result.NotEvaluated)
        AND (FAllTrue.Result = E_Result.NotEvaluated)
        AND (FAllFalse.Result = E_Result.NotEvaluated)
        AND (FContains.Result = E_Result.NotEvaluated);
END_IF;
FActivityMatch := (FEqual.Enabled = FSubjectEnable)
    AND (FEqual.ObservationActive = (FEvaluateSubjects AND FSubjectEnable))
    AND (FEqual.EvaluationActive = (FEvaluateSubjects AND FSubjectEnable))
    AND (FNotEqual.Enabled = FSubjectEnable)
    AND (FNotEqual.ObservationActive = (FEvaluateSubjects AND FSubjectEnable))
    AND (FNotEqual.EvaluationActive = (FEvaluateSubjects AND FSubjectEnable))
    AND (FAllTrue.Enabled = FSubjectEnable)
    AND (FAllTrue.ObservationActive = (FEvaluateSubjects AND FSubjectEnable))
    AND (FAllTrue.EvaluationActive = (FEvaluateSubjects AND FSubjectEnable))
    AND (FAllFalse.Enabled = FSubjectEnable)
    AND (FAllFalse.ObservationActive = (FEvaluateSubjects AND FSubjectEnable))
    AND (FAllFalse.EvaluationActive = (FEvaluateSubjects AND FSubjectEnable))
    AND (FContains.Enabled = FSubjectEnable)
    AND (FContains.ObservationActive = (FEvaluateSubjects AND FSubjectEnable))
    AND (FContains.EvaluationActive = (FEvaluateSubjects AND FSubjectEnable));
END_METHOD

{region 'Documentation'}
(*!
<summary>Initializes outer checks and isolates intentional subject findings.</summary>
*)
{endregion}
METHOD PROTECTED Configure
VAR
    Initialized : BOOL;
END_VAR
FPreparationStateCount := 0;
FTestStateCount := 1;
FResults.Initialize(Parent := THIS^,
    AssertionName := 'Results');
FActivity.Initialize(Parent := THIS^,
    AssertionName := 'Activity');
FInputs.Initialize(Parent := THIS^,
    AssertionName := 'Inputs');
FFindings.Initialize(Parent := THIS^,
    AssertionName := 'Findings');
FSetupValid := FCapture.Initialize(Buffer := FEvents,
    FifoControl := FCaptureFifo,
    Status := FCaptureStatus);
FEqual.BindPublisher(Publisher := FCapture);
Initialized := FEqual.Initialize(Parent := THIS^,
    AssertionName := 'Equal');
FSetupValid := FSetupValid AND Initialized;
FNotEqual.BindPublisher(Publisher := FCapture);
Initialized := FNotEqual.Initialize(Parent := THIS^,
    AssertionName := 'NotEqual');
FSetupValid := FSetupValid AND Initialized;
FAllTrue.BindPublisher(Publisher := FCapture);
Initialized := FAllTrue.Initialize(Parent := THIS^,
    AssertionName := 'AllTrue');
FSetupValid := FSetupValid AND Initialized;
FAllFalse.BindPublisher(Publisher := FCapture);
Initialized := FAllFalse.Initialize(Parent := THIS^,
    AssertionName := 'AllFalse');
FSetupValid := FSetupValid AND Initialized;
FContains.BindPublisher(Publisher := FCapture);
Initialized := FContains.Initialize(Parent := THIS^,
    AssertionName := 'Contains');
FSetupValid := FSetupValid AND Initialized;
END_METHOD

{region 'Documentation'}
(*!
<summary>Completes abort; no asynchronous resource is owned.</summary>
*)
{endregion}
METHOD PROTECTED ProcessAbort
VAR_INPUT
    Enable : BOOL; //! Phase permission supplied by the owning Test Case; FALSE does not authorize progression, while observation may continue.
END_VAR
IF Enable THEN
    CompleteAbort();
END_IF;
END_METHOD

{region 'Documentation'}
(*!
<summary>Latches this call's checks before progression is permitted.</summary>
*)
{endregion}
METHOD PROTECTED ProcessAssertions
VAR_INPUT
    Enable : BOOL; //! Phase permission supplied by the owning Test Case; FALSE does not authorize progression, while observation may continue.
END_VAR
VAR
    Check : BOOL;
END_VAR
Check := Enable AND FObservationReady;
FResults(Enable := Check,
    State := State,
    IN := FResultsMatch);
FActivity(Enable := Check,
    State := State,
    IN := FActivityMatch);
FInputs(Enable := Check,
    State := State,
    IN := FInputsMatch);
FFindings(Enable := Check,
    State := State,
    IN := FFindingsMatch);
IF Check THEN
    FChecked := TRUE;
END_IF;
END_METHOD

{region 'Documentation'}
(*!
<summary>No Preparation phase is needed.</summary>
*)
{endregion}
METHOD PROTECTED ProcessPreparations
VAR_INPUT
    // SA0033: Required hook; this test has no Preparation phase.
    {attribute 'analysis' := '-33'}
    Enable : BOOL; //! Phase permission supplied by the owning Test Case; FALSE does not authorize progression, while observation may continue.
END_VAR
END_METHOD

{region 'Documentation'}
(*!
<summary>Restarts the scenario sequence and outer checks.</summary>
*)
{endregion}
METHOD PROTECTED ProcessReset
FScenario := ScenarioOutsideBitsIgnored;
FChecked := FALSE;
FSubjectEnable := FALSE;
FEvaluateSubjects := FALSE;
FObservationReady := FALSE;
FFirstFailedScenario := 0;
FFailedDuringEvaluation := FALSE;
FCapture.Reset();
ResetSubjects();
FResults.Reset();
FActivity.Reset();
FInputs.Reset();
FFindings.Reset();
CompleteReset();
END_METHOD

{region 'Documentation'}
(*!
<summary>Consumes reset, evaluates, then waits for the outer checks before advancing.</summary>
*)
{endregion}
METHOD PROTECTED ProcessTests
VAR_INPUT
    Enable : BOOL; //! Phase permission supplied by the owning Test Case; FALSE does not authorize progression, while observation may continue.
END_VAR
IF NOT Enable THEN
    RETURN;
END_IF;

IF FChecked THEN
    FChecked := FALSE;
    FObservationReady := FALSE;
    IF FEvaluateSubjects THEN
        IF FScenario = LastScenario THEN
            CompleteTests();
            RETURN;
        END_IF;
        FScenario := FScenario + 1;
    END_IF;
    FEvaluateSubjects := NOT FEvaluateSubjects;
END_IF;

IF NOT SelectScenario() THEN
    RETURN;
END_IF;
FCapture.Reset();
IF NOT FEvaluateSubjects THEN
    ResetSubjects();
END_IF;

CallSubjects();
CheckResults();
CheckInputs();
CheckFindings();
IF (FFirstFailedScenario = 0)
    AND NOT (FResultsMatch AND FActivityMatch AND FInputsMatch AND FFindingsMatch) THEN
    FFirstFailedScenario := FScenario;
    FFailedDuringEvaluation := FEvaluateSubjects;
END_IF;
FObservationReady := TRUE;
END_METHOD

{region 'Documentation'}
(*!
<summary>Queues reset; the next bound FB call consumes it without evaluating.</summary>
*)
{endregion}
METHOD PRIVATE ResetSubjects
FEqual.Reset();
FNotEqual.Reset();
FAllTrue.Reset();
FAllFalse.Reset();
FContains.Reset();
END_METHOD

{region 'Documentation'}
(*!
<summary>Selects explicit stimuli and expected results for one scenario.</summary>
*)
{endregion}
METHOD PRIVATE SelectScenario : BOOL //! TRUE after selecting a supported scenario and its literal expectations; FALSE reports an unknown scenario.
SelectScenario := FALSE;
FSubjectEnable := TRUE;
FWordValue := WORD#16#A505;
FWordMask := WORD#16#00FF;
FExpectedWord := WORD#16#0005;
FWideValue := LWORD#16#8000000000000001;
FWideMask := LWORD#16#8000000000000000;
FForbiddenWide := 0;
FByteValue := BYTE#16#F3;
FByteMask := BYTE#16#03;
FDWordValue := DWORD#16#80000000;
FDWordMask := DWORD#16#00000003;
FContainsValue := LWORD#16#8000000000000000;
FContainsMask := LWORD#16#8000000000000001;
FExpectedBit := TRUE;
CASE FScenario OF
    ScenarioOutsideBitsIgnored:
        FEqualExpectedResult := E_Result.Passed;
        FEqualExpectedFinding := FALSE;
        FNotEqualExpectedResult := E_Result.Passed;
        FNotEqualExpectedFinding := FALSE;
        FAllTrueExpectedResult := E_Result.Passed;
        FAllTrueExpectedFinding := FALSE;
        FAllFalseExpectedResult := E_Result.Passed;
        FAllFalseExpectedFinding := FALSE;
        FContainsExpectedResult := E_Result.Passed;
        FContainsExpectedFinding := FALSE;
    ScenarioPartialSelection:
        FWordValue := WORD#16#A504;
        FWideValue := LWORD#16#0000000000000001;
        FByteValue := BYTE#16#F1;
        FDWordValue := DWORD#16#80000001;
        FEqualExpectedResult := E_Result.Failed;
        FEqualExpectedFinding := TRUE;
        FNotEqualExpectedResult := E_Result.Failed;
        FNotEqualExpectedFinding := TRUE;
        FAllTrueExpectedResult := E_Result.Failed;
        FAllTrueExpectedFinding := TRUE;
        FAllFalseExpectedResult := E_Result.Failed;
        FAllFalseExpectedFinding := TRUE;
        FContainsExpectedResult := E_Result.Passed;
        FContainsExpectedFinding := FALSE;
    ScenarioContainsFalse:
        FExpectedBit := FALSE;
        FEqualExpectedResult := E_Result.Passed;
        FEqualExpectedFinding := FALSE;
        FNotEqualExpectedResult := E_Result.Passed;
        FNotEqualExpectedFinding := FALSE;
        FAllTrueExpectedResult := E_Result.Passed;
        FAllTrueExpectedFinding := FALSE;
        FAllFalseExpectedResult := E_Result.Passed;
        FAllFalseExpectedFinding := FALSE;
        FContainsExpectedResult := E_Result.Passed;
        FContainsExpectedFinding := FALSE;
    ScenarioAllSelectedTrue:
        FContainsValue := LWORD#16#8000000000000001;
        FExpectedBit := FALSE;
        FEqualExpectedResult := E_Result.Passed;
        FEqualExpectedFinding := FALSE;
        FNotEqualExpectedResult := E_Result.Passed;
        FNotEqualExpectedFinding := FALSE;
        FAllTrueExpectedResult := E_Result.Passed;
        FAllTrueExpectedFinding := FALSE;
        FAllFalseExpectedResult := E_Result.Passed;
        FAllFalseExpectedFinding := FALSE;
        FContainsExpectedResult := E_Result.Failed;
        FContainsExpectedFinding := TRUE;
    ScenarioAllSelectedFalse:
        FByteValue := BYTE#16#F0;
        FContainsValue := 0;
        FEqualExpectedResult := E_Result.Passed;
        FEqualExpectedFinding := FALSE;
        FNotEqualExpectedResult := E_Result.Passed;
        FNotEqualExpectedFinding := FALSE;
        FAllTrueExpectedResult := E_Result.Failed;
        FAllTrueExpectedFinding := TRUE;
        FAllFalseExpectedResult := E_Result.Passed;
        FAllFalseExpectedFinding := FALSE;
        FContainsExpectedResult := E_Result.Failed;
        FContainsExpectedFinding := TRUE;
    ScenarioFalsePresent:
        FContainsValue := 0;
        FExpectedBit := FALSE;
        FEqualExpectedResult := E_Result.Passed;
        FEqualExpectedFinding := FALSE;
        FNotEqualExpectedResult := E_Result.Passed;
        FNotEqualExpectedFinding := FALSE;
        FAllTrueExpectedResult := E_Result.Passed;
        FAllTrueExpectedFinding := FALSE;
        FAllFalseExpectedResult := E_Result.Passed;
        FAllFalseExpectedFinding := FALSE;
        FContainsExpectedResult := E_Result.Passed;
        FContainsExpectedFinding := FALSE;
    ScenarioEmptyMasks:
        FWordMask := 0;
        FWideMask := 0;
        FByteMask := 0;
        FDWordMask := 0;
        FContainsMask := 0;
        FEqualExpectedResult := E_Result.Error;
        FEqualExpectedFinding := TRUE;
        FNotEqualExpectedResult := E_Result.Error;
        FNotEqualExpectedFinding := TRUE;
        FAllTrueExpectedResult := E_Result.Error;
        FAllTrueExpectedFinding := TRUE;
        FAllFalseExpectedResult := E_Result.Error;
        FAllFalseExpectedFinding := TRUE;
        FContainsExpectedResult := E_Result.Error;
        FContainsExpectedFinding := TRUE;
ELSE
    Error(Message := 'Unknown variant Assertion scenario.');
    RETURN;
END_CASE;

SelectScenario := TRUE;
END_METHOD

END_FUNCTION_BLOCK

// ---- Framework/Assertions/POU/BasicTypes/LWord/AssertNotEqualMask_LWord.TcPOU
{region 'Documentation'}
(*!
<summary>Checks that selected bits differ from the forbidden masked value.</summary>
*)
{endregion}
FUNCTION_BLOCK AssertNotEqualMask_LWord EXTENDS AssertionBase
VAR_INPUT
    IN : LWORD; //! Actual bitfield.
    Mask : LWORD := 16#FFFFFFFFFFFFFFFF; //! Selects evaluated bits; defaults to all bits. An empty mask produces Error during evaluation.
    Expected : LWORD; //! Forbidden value; bits outside Mask are ignored.
END_VAR

SUPER^();

{region 'Documentation'}
(*!
<summary>Rejects an empty mask before comparing selected bits.</summary>
*)
{endregion}
METHOD PROTECTED Assert
VAR
    Message : STRING(GVL_Constants.MessageLength);
    MaskText : STRING(GVL_Constants.AssertionValueLength);
    ExpectedText : STRING(GVL_Constants.AssertionValueLength);
    ActualText : STRING(GVL_Constants.AssertionValueLength);
END_VAR
VAR CONSTANT
    NoMask : LWORD := 16#00;
    HexDigitCount : USINT := 16;
END_VAR
IF NOT EvaluationActive THEN
    RETURN;
END_IF;

IF Result = E_Result.Error THEN
    RETURN;
END_IF;

IF Mask = NoMask THEN
    MaskText := CreateAssertionTextValue_Hex(Value := Mask,
        DigitCount := HexDigitCount);
    Message := CONCAT('Assertion error: mask must not be empty. Mask = ',
        MaskText);
    Message := CONCAT(Message, '.');
    Error(Message := Message);
    RETURN;
END_IF;

IF Result = E_Result.Failed THEN
    RETURN;
END_IF;

IF (IN AND Mask) = (Expected AND Mask) THEN
    MaskText := CreateAssertionTextValue_Hex(Value := Mask,
        DigitCount := HexDigitCount);
    ExpectedText := CreateAssertionTextValue_Hex(Value := Expected,
        DigitCount := HexDigitCount);
    ActualText := CreateAssertionTextValue_Hex(Value := IN,
        DigitCount := HexDigitCount);
    Message := CONCAT('Assertion failed: selected bits match forbidden value. NotExpected = ',
        ExpectedText);
    Message := CONCAT(Message, ', Mask = ');
    Message := CONCAT(Message, MaskText);
    Message := CONCAT(Message, ', Actual = ');
    Message := CONCAT(Message, ActualText);
    Message := CONCAT(Message, '.');
    Fail(Message := Message);
    RETURN;
END_IF;

Pass();
END_METHOD

END_FUNCTION_BLOCK

// ---- Framework/Assertions/POU/BasicTypes/Byte/AssertTrueMask_Byte.TcPOU
{region 'Documentation'}
(*!
<summary>Checks that all selected bits are TRUE.</summary>
*)
{endregion}
FUNCTION_BLOCK AssertTrueMask_Byte EXTENDS AssertionBase
VAR_INPUT
    IN : BYTE; //! Actual bitfield.
    Mask : BYTE := 16#FF; //! Selects evaluated bits; defaults to all bits. An empty mask produces Error during evaluation.
END_VAR

SUPER^();

{region 'Documentation'}
(*!
<summary>Rejects an empty mask before comparing selected bits.</summary>
*)
{endregion}
METHOD PROTECTED Assert
VAR
    Message : STRING(GVL_Constants.MessageLength);
    MaskText : STRING(GVL_Constants.AssertionValueLength);
    ActualText : STRING(GVL_Constants.AssertionValueLength);
END_VAR
VAR CONSTANT
    NoMask : BYTE := 16#00;
    HexDigitCount : USINT := 2;
END_VAR
IF NOT EvaluationActive THEN
    RETURN;
END_IF;

IF Result = E_Result.Error THEN
    RETURN;
END_IF;

IF Mask = NoMask THEN
    MaskText := CreateAssertionTextValue_Hex(Value := BYTE_TO_LWORD(Mask),
        DigitCount := HexDigitCount);
    Message := CONCAT('Assertion error: mask must not be empty. Mask = ',
        MaskText);
    Message := CONCAT(Message, '.');
    Error(Message := Message);
    RETURN;
END_IF;

IF Result = E_Result.Failed THEN
    RETURN;
END_IF;

IF (IN AND Mask) <> Mask THEN
    MaskText := CreateAssertionTextValue_Hex(Value := BYTE_TO_LWORD(Mask),
        DigitCount := HexDigitCount);
    ActualText := CreateAssertionTextValue_Hex(Value := BYTE_TO_LWORD(IN),
        DigitCount := HexDigitCount);
    Message := CONCAT('Assertion failed: selected bits are not all TRUE. Mask = ',
        MaskText);
    Message := CONCAT(Message, ', Actual = ');
    Message := CONCAT(Message, ActualText);
    Message := CONCAT(Message, '.');
    Fail(Message := Message);
    RETURN;
END_IF;

Pass();
END_METHOD

END_FUNCTION_BLOCK

// ---- Framework/Assertions/POU/BasicTypes/DWord/AssertFalseMask_DWord.TcPOU
{region 'Documentation'}
(*!
<summary>Checks that all selected bits are FALSE.</summary>
*)
{endregion}
FUNCTION_BLOCK AssertFalseMask_DWord EXTENDS AssertionBase
VAR_INPUT
    IN : DWORD; //! Actual bitfield.
    Mask : DWORD := 16#FFFFFFFF; //! Selects evaluated bits; defaults to all bits. An empty mask produces Error during evaluation.
END_VAR

SUPER^();

{region 'Documentation'}
(*!
<summary>Rejects an empty mask before comparing selected bits.</summary>
*)
{endregion}
METHOD PROTECTED Assert
VAR
    Message : STRING(GVL_Constants.MessageLength);
    MaskText : STRING(GVL_Constants.AssertionValueLength);
    ActualText : STRING(GVL_Constants.AssertionValueLength);
END_VAR
VAR CONSTANT
    NoMask : DWORD := 16#00;
    HexDigitCount : USINT := 8;
END_VAR
IF NOT EvaluationActive THEN
    RETURN;
END_IF;

IF Result = E_Result.Error THEN
    RETURN;
END_IF;

IF Mask = NoMask THEN
    MaskText := CreateAssertionTextValue_Hex(Value := DWORD_TO_LWORD(Mask),
        DigitCount := HexDigitCount);
    Message := CONCAT('Assertion error: mask must not be empty. Mask = ',
        MaskText);
    Message := CONCAT(Message, '.');
    Error(Message := Message);
    RETURN;
END_IF;

IF Result = E_Result.Failed THEN
    RETURN;
END_IF;

IF (IN AND Mask) <> NoMask THEN
    MaskText := CreateAssertionTextValue_Hex(Value := DWORD_TO_LWORD(Mask),
        DigitCount := HexDigitCount);
    ActualText := CreateAssertionTextValue_Hex(Value := DWORD_TO_LWORD(IN),
        DigitCount := HexDigitCount);
    Message := CONCAT('Assertion failed: selected bits are not all FALSE. Mask = ',
        MaskText);
    Message := CONCAT(Message, ', Actual = ');
    Message := CONCAT(Message, ActualText);
    Message := CONCAT(Message, '.');
    Fail(Message := Message);
    RETURN;
END_IF;

Pass();
END_METHOD

END_FUNCTION_BLOCK

// ---- Framework/Assertions/POU/BasicTypes/LWord/AssertContainsBit_LWord.TcPOU
{region 'Documentation'}
(*!
<summary>Checks that at least one selected bit equals the expected Boolean value.</summary>
*)
{endregion}
FUNCTION_BLOCK AssertContainsBit_LWord EXTENDS AssertionBase
VAR_INPUT
    IN : LWORD; //! Actual bitfield.
    Mask : LWORD := 16#FFFFFFFFFFFFFFFF; //! Selects evaluated bits; defaults to all bits. An empty mask produces Error during evaluation.
    Expected : BOOL; //! Expected value of at least one selected bit.
END_VAR

SUPER^();

{region 'Documentation'}
(*!
<summary>Rejects an empty mask before checking for a matching selected bit.</summary>
*)
{endregion}
METHOD PROTECTED Assert
VAR
    ContainsBit : BOOL;
    Message : STRING(GVL_Constants.MessageLength);
    MaskText : STRING(GVL_Constants.AssertionValueLength);
    ActualText : STRING(GVL_Constants.AssertionValueLength);
END_VAR
VAR CONSTANT
    NoMask : LWORD := 16#00;
    HexDigitCount : USINT := 16;
END_VAR
IF NOT EvaluationActive THEN
    RETURN;
END_IF;

IF Result = E_Result.Error THEN
    RETURN;
END_IF;

IF Mask = NoMask THEN
    MaskText := CreateAssertionTextValue_Hex(Value := Mask,
        DigitCount := HexDigitCount);
    Message := CONCAT('Assertion error: mask must not be empty. Mask = ',
        MaskText);
    Message := CONCAT(Message, '.');
    Error(Message := Message);
    RETURN;
END_IF;

IF Result = E_Result.Failed THEN
    RETURN;
END_IF;

IF Expected THEN
    ContainsBit := (IN AND Mask) <> NoMask;
ELSE
    ContainsBit := (IN AND Mask) <> Mask;
END_IF;

IF NOT ContainsBit THEN
    MaskText := CreateAssertionTextValue_Hex(Value := Mask,
        DigitCount := HexDigitCount);
    ActualText := CreateAssertionTextValue_Hex(Value := IN,
        DigitCount := HexDigitCount);
    Message := CONCAT('Assertion failed: selected bits do not contain expected bit value. Expected = ',
        BOOL_TO_STRING(Expected));
    Message := CONCAT(Message, ', Mask = ');
    Message := CONCAT(Message, MaskText);
    Message := CONCAT(Message, ', Actual = ');
    Message := CONCAT(Message, ActualText);
    Message := CONCAT(Message, '.');
    Fail(Message := Message);
    RETURN;
END_IF;

Pass();
END_METHOD

END_FUNCTION_BLOCK

// ---- SelfTests/TestCases/TestSuite_AssertionVariants/Test_AssertionCountPredicates.TcPOU
{region 'Documentation'}
(*!
<summary>Checks residual count and length relations around the known value two.</summary>
<description>
Each independent scenario consumes a bound reset, a baseline and three edge samples before evaluation.
ProcessAssertions checks the observation before ProcessTests advances.
SelectScenario holds explicit expected results; no production algorithm is mirrored.
Expected findings remain in the local capture; only outer checks affect the test result.
FirstFailedScenario and FailedDuringEvaluation retain the first mismatch.
Each scenario resets, observes two rising/falling edges, then evaluates once. Array fixtures contain two tokens and a two-element prefix; search algorithms are not reproduced.
</description>
*)
{endregion}
FUNCTION_BLOCK Test_AssertionCountPredicates EXTENDS TestCaseBase
VAR
    FRising : AssertRisingEdgeCntGreaterThan;
    FRisingExpectedResult : E_Result;
    FRisingExpectedFinding : BOOL;
    FFalling : AssertFallingEdgeCntLessEqual;
    FFallingExpectedResult : E_Result;
    FFallingExpectedFinding : BOOL;
    FValueCount : AssertValueTokenCntNotEqual_Byte;
    FValueCountExpectedResult : E_Result;
    FValueCountExpectedFinding : BOOL;
    FOutsideCount : AssertArrayTokenCntNotInRange_Word;
    FOutsideCountExpectedResult : E_Result;
    FOutsideCountExpectedFinding : BOOL;
    FBelowCount : AssertArrayTokenCntLessThan_Byte;
    FBelowCountExpectedResult : E_Result;
    FBelowCountExpectedFinding : BOOL;
    FPrefixLength : AssertLengthUntilArrayGreaterEqual_Word;
    FPrefixLengthExpectedResult : E_Result;
    FPrefixLengthExpectedFinding : BOOL;
    FData : ARRAY[1..6] OF BYTE;
    FDataBefore : ARRAY[1..6] OF BYTE;
    FWideData : ARRAY[1..6] OF WORD;
    FWideDataBefore : ARRAY[1..6] OF WORD;
    FToken : ARRAY[4..5] OF BYTE;
    FTokenBefore : ARRAY[4..5] OF BYTE;
    FWideToken : ARRAY[-2..-1] OF WORD;
    FWideTokenBefore : ARRAY[-2..-1] OF WORD;
    FPhase : UINT;
    FSample : BOOL;
    FLimit : UINT;
    FRangeMinimum : UINT;
    FRangeMaximum : UINT;
    FSubjectEnable : BOOL;
    FCapture : EventBuffer;
    FEvents : ARRAY[1..CaptureLength] OF ST_Event;
    FCaptureFifo : ST_FifoStatus;
    FCaptureStatus : ST_EventBufferStatus;
    FSetupValid : BOOL;
    FScenario : UINT;
    FChecked : BOOL;
    FEvaluateSubjects : BOOL;
    FObservationReady : BOOL;
    FFirstFailedScenario : UINT;
    FFailedDuringEvaluation : BOOL;
    FResultsMatch : BOOL;
    FResults : AssertTrue;
    FActivityMatch : BOOL;
    FActivity : AssertTrue;
    FInputsMatch : BOOL;
    FInputs : AssertTrue;
    FFindingsMatch : BOOL;
    FFindings : AssertTrue;
END_VAR
VAR CONSTANT
    CaptureLength : UINT := 12;
    PhaseReset : UINT := 0;
    PhaseBaseline : UINT := 1;
    PhaseFirstEdge : UINT := 2;
    PhaseOppositeEdge : UINT := 3;
    PhaseSecondEdge : UINT := 4;
    PhaseEvaluate : UINT := 5;
    ScenarioBelowCount : UINT := 1;
    ScenarioEqualCount : UINT := 2;
    ScenarioAboveCount : UINT := 3;
    ScenarioInclusiveLower : UINT := 4;
    ScenarioInclusiveUpper : UINT := 5;
    ScenarioReversedBounds : UINT := 6;
    LastScenario : UINT := ScenarioReversedBounds;
END_VAR

SUPER^();

{region 'Documentation'}
(*!
<summary>Aggregates only outer checks, not intentionally failing subjects.</summary>
*)
{endregion}
METHOD PROTECTED AggregateResults
VAR_INPUT
    Aggregator : I_ResultAggregator; //! Borrowed result sink owned by the outer Test Case; add this test's checking Assertions without resetting or retaining the sink.
END_VAR
Aggregator.AddProvider(Provider := FResults);
Aggregator.AddProvider(Provider := FActivity);
Aggregator.AddProvider(Provider := FInputs);
Aggregator.AddProvider(Provider := FFindings);
END_METHOD

{region 'Documentation'}
(*!
<summary>Calls each inherited production subject once with caller-owned input storage.</summary>
*)
{endregion}
METHOD PRIVATE CallSubjects
FRising(Enable := FSubjectEnable,
    Evaluate := FEvaluateSubjects,
    State := E_State.Running,
    IN := FSample,
    Minimum := FLimit);
FFalling(Enable := FSubjectEnable,
    Evaluate := FEvaluateSubjects,
    State := E_State.Running,
    IN := NOT FSample,
    Maximum := FLimit);
FValueCount(Enable := FEvaluateSubjects,
    State := E_State.Running,
    StartIndex := 1,
    Length := 6,
    Expected := FLimit,
    Token := 1,
    IN := FData);
FOutsideCount(Enable := FEvaluateSubjects,
    State := E_State.Running,
    StartIndex := 1,
    Length := 6,
    Minimum := FRangeMinimum,
    Maximum := FRangeMaximum,
    IN := FWideData,
    Token := FWideToken);
FBelowCount(Enable := FEvaluateSubjects,
    State := E_State.Running,
    StartIndex := 1,
    Length := 6,
    Maximum := FLimit,
    IN := FData,
    Token := FToken);
FPrefixLength(Enable := FEvaluateSubjects,
    State := E_State.Running,
    StartIndex := 1,
    Length := 6,
    Expected := UINT_TO_USINT(FLimit),
    IN := FWideData,
    Token := FWideToken);
END_METHOD

{region 'Documentation'}
(*!
<summary>Checks one subject finding in call order; expected outcomes come from the scenario.</summary>
*)
{endregion}
METHOD PRIVATE CheckFinding : BOOL //! TRUE when the required finding checks pass; calls requiring no finding also succeed.
VAR_INPUT
    Subject : I_Assertion; //! Assertion interface supplying the expected finding identity.
    ExpectedResult : E_Result; //! Independently authored result expected in the captured finding.
    ExpectedFinding : BOOL; //! TRUE when this scenario requires a finding during active evaluation.
END_VAR
VAR_IN_OUT
    Index : UINT; //! One-based next finding index; advanced when this call checks a required finding.
END_VAR
CheckFinding := TRUE;
IF FEvaluateSubjects AND ExpectedFinding THEN
    CheckFinding := (FEvents[Index].SequenceId = UINT_TO_UDINT(Index))
        AND (FEvents[Index].Name = Subject.Name)
        AND (FEvents[Index].OwnerScope = E_OwnerScope.Assertion)
        AND (FEvents[Index].EventType = E_EventType.Result)
        AND (FEvents[Index].State = E_State.Running)
        AND (FEvents[Index].Result = ExpectedResult)
        AND (FEvents[Index].Message <> '');
    Index := Index + 1;
END_IF;
END_METHOD

{region 'Documentation'}
(*!
<summary>Checks exact finding count and identities; at most one finding per subject.</summary>
*)
{endregion}
METHOD PRIVATE CheckFindings
VAR
    Index : UINT;
    Matches : BOOL;
END_VAR
Index := 1;
FFindingsMatch := TRUE;
Matches := CheckFinding(Subject := FRising,
    ExpectedResult := FRisingExpectedResult,
    ExpectedFinding := FRisingExpectedFinding,
    Index := Index);
FFindingsMatch := FFindingsMatch AND Matches;
Matches := CheckFinding(Subject := FFalling,
    ExpectedResult := FFallingExpectedResult,
    ExpectedFinding := FFallingExpectedFinding,
    Index := Index);
FFindingsMatch := FFindingsMatch AND Matches;
Matches := CheckFinding(Subject := FValueCount,
    ExpectedResult := FValueCountExpectedResult,
    ExpectedFinding := FValueCountExpectedFinding,
    Index := Index);
FFindingsMatch := FFindingsMatch AND Matches;
Matches := CheckFinding(Subject := FOutsideCount,
    ExpectedResult := FOutsideCountExpectedResult,
    ExpectedFinding := FOutsideCountExpectedFinding,
    Index := Index);
FFindingsMatch := FFindingsMatch AND Matches;
Matches := CheckFinding(Subject := FBelowCount,
    ExpectedResult := FBelowCountExpectedResult,
    ExpectedFinding := FBelowCountExpectedFinding,
    Index := Index);
FFindingsMatch := FFindingsMatch AND Matches;
Matches := CheckFinding(Subject := FPrefixLength,
    ExpectedResult := FPrefixLengthExpectedResult,
    ExpectedFinding := FPrefixLengthExpectedFinding,
    Index := Index);
FFindingsMatch := FFindingsMatch AND Matches;
FFindingsMatch := FFindingsMatch
    AND (FCaptureStatus.SequenceId = UINT_TO_UDINT(Index - 1))
    AND (FCaptureStatus.LostEventCount = 0);
IF FEvaluateSubjects AND (FScenario = ScenarioBelowCount) THEN
    // SA0175: Fixed byte-substring checks of bounded diagnostic messages; no character offsets.
    {analysis -175}
    FFindingsMatch := FFindingsMatch
        AND (FIND(FEvents[1].Message, 'Maximum = 1') > 0)
        AND (FIND(FEvents[1].Message, 'Actual = 2') > 0)
        AND (FIND(FEvents[2].Message, 'Maximum = 1') > 0)
        AND (FIND(FEvents[2].Message, 'Actual = 2') > 0);
    {analysis +175}
END_IF;
IF FEvaluateSubjects AND (FScenario = ScenarioAboveCount) THEN
    // SA0175: Fixed byte-substring checks of bounded diagnostic messages; no character offsets.
    {analysis -175}
    FFindingsMatch := FFindingsMatch
        AND (FIND(FEvents[1].Message, 'Minimum = 3') > 0)
        AND (FIND(FEvents[1].Message, 'Actual = 2') > 0)
        AND (FIND(FEvents[2].Message, 'Expected = 3') > 0)
        AND (FIND(FEvents[2].Message, 'Actual = 2') > 0);
    {analysis +175}
END_IF;
END_METHOD

{region 'Documentation'}
(*!
<summary>Rejects incomplete subject, capture or outer Assertion setup.</summary>
*)
{endregion}
METHOD PROTECTED CheckInitialization : BOOL //! TRUE when the inherited initialization check and this concrete fixture check both accept the setup.
CheckInitialization := SUPER^.CheckInitialization();
IF NOT CheckInitialization THEN
    RETURN;
END_IF;

CheckInitialization := FSetupValid
    AND FResults.IsInitialized
    AND FActivity.IsInitialized
    AND FInputs.IsInitialized
    AND FFindings.IsInitialized;
IF NOT CheckInitialization THEN
    EventPublisher.PublishEvent(Event := CreateFrameworkEvent(Name := Name,
        ResourceName := '',
        State := State,
        Severity := E_EventSeverity.Error,
        Message := 'Variant selftest setup failed.'));
END_IF;
END_METHOD

{region 'Documentation'}
(*!
<summary>Verifies input preservation without using the tested comparison algorithm.</summary>
*)
{endregion}
METHOD PRIVATE CheckInputs
VAR
    Index : DINT;
END_VAR
FInputsMatch := TRUE;
FOR Index := 1 TO 6 DO
    FInputsMatch := FInputsMatch AND (FData[Index] = FDataBefore[Index]);
END_FOR;
FOR Index := 1 TO 6 DO
    FInputsMatch := FInputsMatch AND (FWideData[Index] = FWideDataBefore[Index]);
END_FOR;
FOR Index := 4 TO 5 DO
    FInputsMatch := FInputsMatch AND (FToken[Index] = FTokenBefore[Index]);
END_FOR;
FOR Index := -2 TO -1 DO
    FInputsMatch := FInputsMatch AND (FWideToken[Index] = FWideTokenBefore[Index]);
END_FOR;
END_METHOD

{region 'Documentation'}
(*!
<summary>Checks literal evaluation results, or NotEvaluated while building the known count.</summary>
*)
{endregion}
METHOD PRIVATE CheckResults
VAR
    ExpectedEdgeCount : UINT;
    ExpectedArrayCount : UINT;
    ExpectedOutsideCount : UINT;
END_VAR
IF FEvaluateSubjects THEN
    FResultsMatch := (FRising.Result = FRisingExpectedResult)
        AND (FFalling.Result = FFallingExpectedResult)
        AND (FValueCount.Result = FValueCountExpectedResult)
        AND (FOutsideCount.Result = FOutsideCountExpectedResult)
        AND (FBelowCount.Result = FBelowCountExpectedResult)
        AND (FPrefixLength.Result = FPrefixLengthExpectedResult);
ELSE
    FResultsMatch := (FRising.Result = E_Result.NotEvaluated)
        AND (FFalling.Result = E_Result.NotEvaluated)
        AND (FValueCount.Result = E_Result.NotEvaluated)
        AND (FOutsideCount.Result = E_Result.NotEvaluated)
        AND (FBelowCount.Result = E_Result.NotEvaluated)
        AND (FPrefixLength.Result = E_Result.NotEvaluated);
END_IF;
FActivityMatch := (FRising.Enabled = FSubjectEnable)
    AND (FRising.ObservationActive = FSubjectEnable)
    AND (FRising.EvaluationActive = FEvaluateSubjects)
    AND (FFalling.Enabled = FSubjectEnable)
    AND (FFalling.ObservationActive = FSubjectEnable)
    AND (FFalling.EvaluationActive = FEvaluateSubjects)
    AND (FValueCount.Enabled = FEvaluateSubjects)
    AND (FValueCount.EvaluationActive = FEvaluateSubjects)
    AND (FOutsideCount.Enabled = FEvaluateSubjects)
    AND (FOutsideCount.EvaluationActive = FEvaluateSubjects)
    AND (FBelowCount.Enabled = FEvaluateSubjects)
    AND (FBelowCount.EvaluationActive = FEvaluateSubjects)
    AND (FPrefixLength.Enabled = FEvaluateSubjects)
    AND (FPrefixLength.EvaluationActive = FEvaluateSubjects);
ExpectedEdgeCount := 0;
IF (FPhase = PhaseFirstEdge) OR (FPhase = PhaseOppositeEdge) THEN
    ExpectedEdgeCount := 1;
ELSIF (FPhase = PhaseSecondEdge) OR (FPhase = PhaseEvaluate) THEN
    ExpectedEdgeCount := 2;
END_IF;
ExpectedArrayCount := 0;
ExpectedOutsideCount := 0;
IF FEvaluateSubjects THEN
    ExpectedArrayCount := 2;
    IF FScenario <> ScenarioReversedBounds THEN
        ExpectedOutsideCount := 2;
    END_IF;
END_IF;
FResultsMatch := FResultsMatch
    AND (FRising.EdgeCount = ExpectedEdgeCount)
    AND (FFalling.EdgeCount = ExpectedEdgeCount)
    AND (FValueCount.TokenCount = ExpectedArrayCount)
    AND (FOutsideCount.TokenCount = ExpectedOutsideCount)
    AND (FBelowCount.TokenCount = ExpectedArrayCount);
END_METHOD

{region 'Documentation'}
(*!
<summary>Initializes outer checks and isolates intentional subject findings.</summary>
*)
{endregion}
METHOD PROTECTED Configure
VAR
    Initialized : BOOL;
END_VAR
FPreparationStateCount := 0;
FTestStateCount := 1;
FResults.Initialize(Parent := THIS^,
    AssertionName := 'Results');
FActivity.Initialize(Parent := THIS^,
    AssertionName := 'Activity');
FInputs.Initialize(Parent := THIS^,
    AssertionName := 'Inputs');
FFindings.Initialize(Parent := THIS^,
    AssertionName := 'Findings');
FSetupValid := FCapture.Initialize(Buffer := FEvents,
    FifoControl := FCaptureFifo,
    Status := FCaptureStatus);
FRising.BindPublisher(Publisher := FCapture);
Initialized := FRising.Initialize(Parent := THIS^,
    AssertionName := 'Rising');
FSetupValid := FSetupValid AND Initialized;
FFalling.BindPublisher(Publisher := FCapture);
Initialized := FFalling.Initialize(Parent := THIS^,
    AssertionName := 'Falling');
FSetupValid := FSetupValid AND Initialized;
FValueCount.BindPublisher(Publisher := FCapture);
Initialized := FValueCount.Initialize(Parent := THIS^,
    AssertionName := 'ValueCount');
FSetupValid := FSetupValid AND Initialized;
FOutsideCount.BindPublisher(Publisher := FCapture);
Initialized := FOutsideCount.Initialize(Parent := THIS^,
    AssertionName := 'OutsideCount');
FSetupValid := FSetupValid AND Initialized;
FBelowCount.BindPublisher(Publisher := FCapture);
Initialized := FBelowCount.Initialize(Parent := THIS^,
    AssertionName := 'BelowCount');
FSetupValid := FSetupValid AND Initialized;
FPrefixLength.BindPublisher(Publisher := FCapture);
Initialized := FPrefixLength.Initialize(Parent := THIS^,
    AssertionName := 'PrefixLength');
FSetupValid := FSetupValid AND Initialized;
END_METHOD

{region 'Documentation'}
(*!
<summary>Completes abort; no asynchronous resource is owned.</summary>
*)
{endregion}
METHOD PROTECTED ProcessAbort
VAR_INPUT
    Enable : BOOL; //! Phase permission supplied by the owning Test Case; FALSE does not authorize progression, while observation may continue.
END_VAR
IF Enable THEN
    CompleteAbort();
END_IF;
END_METHOD

{region 'Documentation'}
(*!
<summary>Latches this call's checks before progression is permitted.</summary>
*)
{endregion}
METHOD PROTECTED ProcessAssertions
VAR_INPUT
    Enable : BOOL; //! Phase permission supplied by the owning Test Case; FALSE does not authorize progression, while observation may continue.
END_VAR
VAR
    Check : BOOL;
END_VAR
Check := Enable AND FObservationReady;
FResults(Enable := Check,
    State := State,
    IN := FResultsMatch);
FActivity(Enable := Check,
    State := State,
    IN := FActivityMatch);
FInputs(Enable := Check,
    State := State,
    IN := FInputsMatch);
FFindings(Enable := Check,
    State := State,
    IN := FFindingsMatch);
IF Check THEN
    FChecked := TRUE;
END_IF;
END_METHOD

{region 'Documentation'}
(*!
<summary>No Preparation phase is needed.</summary>
*)
{endregion}
METHOD PROTECTED ProcessPreparations
VAR_INPUT
    // SA0033: Required hook; this test has no Preparation phase.
    {attribute 'analysis' := '-33'}
    Enable : BOOL; //! Phase permission supplied by the owning Test Case; FALSE does not authorize progression, while observation may continue.
END_VAR
END_METHOD

{region 'Documentation'}
(*!
<summary>Restarts the scenario sequence and outer checks.</summary>
*)
{endregion}
METHOD PROTECTED ProcessReset
FScenario := ScenarioBelowCount;
FPhase := PhaseReset;
FChecked := FALSE;
FSubjectEnable := FALSE;
FEvaluateSubjects := FALSE;
FObservationReady := FALSE;
FFirstFailedScenario := 0;
FFailedDuringEvaluation := FALSE;
FCapture.Reset();
ResetSubjects();
FResults.Reset();
FActivity.Reset();
FInputs.Reset();
FFindings.Reset();
CompleteReset();
END_METHOD

{region 'Documentation'}
(*!
<summary>Builds a known count over successive PLC cycles, then evaluates one relation boundary.</summary>
*)
{endregion}
METHOD PROTECTED ProcessTests
VAR_INPUT
    Enable : BOOL; //! Phase permission supplied by the owning Test Case; FALSE does not authorize progression, while observation may continue.
END_VAR
IF NOT Enable THEN
    RETURN;
END_IF;

IF FChecked THEN
    FChecked := FALSE;
    FObservationReady := FALSE;
    IF FPhase = PhaseEvaluate THEN
        IF FScenario = LastScenario THEN
            CompleteTests();
            RETURN;
        END_IF;
        FScenario := FScenario + 1;
        FPhase := PhaseReset;
    ELSE
        FPhase := FPhase + 1;
    END_IF;
END_IF;

IF NOT SelectScenario() THEN
    RETURN;
END_IF;
FSubjectEnable := (FPhase >= PhaseBaseline) AND (FPhase <= PhaseSecondEdge);
FEvaluateSubjects := FPhase = PhaseEvaluate;
FSample := (FPhase = PhaseFirstEdge) OR (FPhase = PhaseSecondEdge);
FCapture.Reset();
IF FPhase = PhaseReset THEN
    ResetSubjects();
END_IF;
FDataBefore := FData;
FWideDataBefore := FWideData;
FTokenBefore := FToken;
FWideTokenBefore := FWideToken;
CallSubjects();
CheckResults();
CheckInputs();
CheckFindings();
IF (FFirstFailedScenario = 0)
    AND NOT (FResultsMatch AND FActivityMatch AND FInputsMatch AND FFindingsMatch) THEN
    FFirstFailedScenario := FScenario;
    FFailedDuringEvaluation := FEvaluateSubjects;
END_IF;
FObservationReady := TRUE;
END_METHOD

{region 'Documentation'}
(*!
<summary>Queues reset; the next bound FB call consumes it without evaluating.</summary>
*)
{endregion}
METHOD PRIVATE ResetSubjects
FRising.Reset();
FFalling.Reset();
FValueCount.Reset();
FOutsideCount.Reset();
FBelowCount.Reset();
FPrefixLength.Reset();
END_METHOD

{region 'Documentation'}
(*!
<summary>Selects explicit stimuli and expected results for one scenario.</summary>
*)
{endregion}
METHOD PRIVATE SelectScenario : BOOL //! TRUE after selecting a supported scenario and its literal expectations; FALSE reports an unknown scenario.
SelectScenario := FALSE;
FSubjectEnable := TRUE;
FData[1] := 9;
FData[2] := 9;
FData[3] := 1;
FData[4] := 2;
FData[5] := 1;
FData[6] := 2;
FWideData[1] := 9;
FWideData[2] := 9;
FWideData[3] := WORD#16#0101;
FWideData[4] := WORD#16#0202;
FWideData[5] := WORD#16#0101;
FWideData[6] := WORD#16#0202;
FToken[4] := 1;
FToken[5] := 2;
FWideToken[-2] := WORD#16#0101;
FWideToken[-1] := WORD#16#0202;
FLimit := 2;
FRangeMinimum := 2;
FRangeMaximum := 2;
CASE FScenario OF
    ScenarioBelowCount:
        FLimit := 1;
        FRangeMinimum := 1;
        FRangeMaximum := 1;
        FRisingExpectedResult := E_Result.Passed;
        FRisingExpectedFinding := FALSE;
        FFallingExpectedResult := E_Result.Failed;
        FFallingExpectedFinding := TRUE;
        FValueCountExpectedResult := E_Result.Passed;
        FValueCountExpectedFinding := FALSE;
        FOutsideCountExpectedResult := E_Result.Passed;
        FOutsideCountExpectedFinding := FALSE;
        FBelowCountExpectedResult := E_Result.Failed;
        FBelowCountExpectedFinding := TRUE;
        FPrefixLengthExpectedResult := E_Result.Passed;
        FPrefixLengthExpectedFinding := FALSE;
    ScenarioEqualCount:
        FRisingExpectedResult := E_Result.Failed;
        FRisingExpectedFinding := TRUE;
        FFallingExpectedResult := E_Result.Passed;
        FFallingExpectedFinding := FALSE;
        FValueCountExpectedResult := E_Result.Failed;
        FValueCountExpectedFinding := TRUE;
        FOutsideCountExpectedResult := E_Result.Failed;
        FOutsideCountExpectedFinding := TRUE;
        FBelowCountExpectedResult := E_Result.Failed;
        FBelowCountExpectedFinding := TRUE;
        FPrefixLengthExpectedResult := E_Result.Passed;
        FPrefixLengthExpectedFinding := FALSE;
    ScenarioAboveCount:
        FLimit := 3;
        FRangeMinimum := 3;
        FRangeMaximum := 3;
        FRisingExpectedResult := E_Result.Failed;
        FRisingExpectedFinding := TRUE;
        FFallingExpectedResult := E_Result.Passed;
        FFallingExpectedFinding := FALSE;
        FValueCountExpectedResult := E_Result.Passed;
        FValueCountExpectedFinding := FALSE;
        FOutsideCountExpectedResult := E_Result.Passed;
        FOutsideCountExpectedFinding := FALSE;
        FBelowCountExpectedResult := E_Result.Passed;
        FBelowCountExpectedFinding := FALSE;
        FPrefixLengthExpectedResult := E_Result.Failed;
        FPrefixLengthExpectedFinding := TRUE;
    ScenarioInclusiveLower:
        FRangeMinimum := 2;
        FRangeMaximum := 3;
        FRisingExpectedResult := E_Result.Failed;
        FRisingExpectedFinding := TRUE;
        FFallingExpectedResult := E_Result.Passed;
        FFallingExpectedFinding := FALSE;
        FValueCountExpectedResult := E_Result.Failed;
        FValueCountExpectedFinding := TRUE;
        FOutsideCountExpectedResult := E_Result.Failed;
        FOutsideCountExpectedFinding := TRUE;
        FBelowCountExpectedResult := E_Result.Failed;
        FBelowCountExpectedFinding := TRUE;
        FPrefixLengthExpectedResult := E_Result.Passed;
        FPrefixLengthExpectedFinding := FALSE;
    ScenarioInclusiveUpper:
        FRangeMinimum := 1;
        FRangeMaximum := 2;
        FRisingExpectedResult := E_Result.Failed;
        FRisingExpectedFinding := TRUE;
        FFallingExpectedResult := E_Result.Passed;
        FFallingExpectedFinding := FALSE;
        FValueCountExpectedResult := E_Result.Failed;
        FValueCountExpectedFinding := TRUE;
        FOutsideCountExpectedResult := E_Result.Failed;
        FOutsideCountExpectedFinding := TRUE;
        FBelowCountExpectedResult := E_Result.Failed;
        FBelowCountExpectedFinding := TRUE;
        FPrefixLengthExpectedResult := E_Result.Passed;
        FPrefixLengthExpectedFinding := FALSE;
    ScenarioReversedBounds:
        FRangeMinimum := 3;
        FRangeMaximum := 1;
        FRisingExpectedResult := E_Result.Failed;
        FRisingExpectedFinding := TRUE;
        FFallingExpectedResult := E_Result.Passed;
        FFallingExpectedFinding := FALSE;
        FValueCountExpectedResult := E_Result.Failed;
        FValueCountExpectedFinding := TRUE;
        FOutsideCountExpectedResult := E_Result.Error;
        FOutsideCountExpectedFinding := TRUE;
        FBelowCountExpectedResult := E_Result.Failed;
        FBelowCountExpectedFinding := TRUE;
        FPrefixLengthExpectedResult := E_Result.Passed;
        FPrefixLengthExpectedFinding := FALSE;
ELSE
    Error(Message := 'Unknown variant Assertion scenario.');
    RETURN;
END_CASE;

SelectScenario := TRUE;
END_METHOD

END_FUNCTION_BLOCK

// ---- SelfTests/TestCases/TestSuite_AssertionVariants/Test_AssertionNarrowIntegers.TcPOU
{region 'Documentation'}
(*!
<summary>Checks narrow integers with isolated production subjects.</summary>
<description>
Each independent scenario consumes a bound reset call before its evaluation call.
ProcessAssertions checks the observation before ProcessTests advances.
SelectScenario holds explicit expected results; no production algorithm is mirrored.
Expected findings remain in the local capture; only outer checks affect the test result.
FirstFailedScenario and FailedDuringEvaluation retain the first mismatch.
Each scenario uses literal typed inputs at the declared operand widths.
</description>
*)
{endregion}
FUNCTION_BLOCK Test_AssertionNarrowIntegers EXTENDS TestCaseBase
VAR
    FSigned : AssertGreaterThan_SInt;
    FSignedExpectedResult : E_Result;
    FSignedExpectedFinding : BOOL;
    FUnsigned : AssertInRange_USInt;
    FUnsignedExpectedResult : E_Result;
    FUnsignedExpectedFinding : BOOL;

    FSignedValue : SINT;
    FSignedMinimum : SINT;
    FUnsignedValue : USINT;
    FUnsignedMinimum : USINT;
    FUnsignedMaximum : USINT;
    FSubjectEnable : BOOL;
    FCapture : EventBuffer;
    FEvents : ARRAY[1..CaptureLength] OF ST_Event;
    FCaptureFifo : ST_FifoStatus;
    FCaptureStatus : ST_EventBufferStatus;
    FSetupValid : BOOL;
    FScenario : UINT;
    FChecked : BOOL;
    FEvaluateSubjects : BOOL;
    FObservationReady : BOOL;
    FFirstFailedScenario : UINT;
    FFailedDuringEvaluation : BOOL;
    FResultsMatch : BOOL;
    FResults : AssertTrue;
    FActivityMatch : BOOL;
    FActivity : AssertTrue;
    FInputsMatch : BOOL;
    FInputs : AssertTrue;
    FFindingsMatch : BOOL;
    FFindings : AssertTrue;
END_VAR
VAR CONSTANT
    CaptureLength : UINT := 8;
    ScenarioLowerLimits : UINT := 1;
    ScenarioUpperLimits : UINT := 2;
    ScenarioEqualSignedMinimum : UINT := 3;
    ScenarioOutsideRange : UINT := 4;
    ScenarioAboveMaximum : UINT := 5;
    ScenarioSingleValue : UINT := 6;
    ScenarioReversedRange : UINT := 7;
    LastScenario : UINT := ScenarioReversedRange;
END_VAR

SUPER^();

{region 'Documentation'}
(*!
<summary>Aggregates only outer checks, not intentionally failing subjects.</summary>
*)
{endregion}
METHOD PROTECTED AggregateResults
VAR_INPUT
    Aggregator : I_ResultAggregator; //! Borrowed result sink owned by the outer Test Case; add this test's checking Assertions without resetting or retaining the sink.
END_VAR
Aggregator.AddProvider(Provider := FResults);
Aggregator.AddProvider(Provider := FActivity);
Aggregator.AddProvider(Provider := FInputs);
Aggregator.AddProvider(Provider := FFindings);
END_METHOD

{region 'Documentation'}
(*!
<summary>Calls each inherited production subject once with caller-owned input storage.</summary>
*)
{endregion}
METHOD PRIVATE CallSubjects
FSigned(Enable := FSubjectEnable,
    State := E_State.Running,
    IN := FSignedValue,
    Minimum := FSignedMinimum);
FUnsigned(Enable := FSubjectEnable,
    State := E_State.Running,
    IN := FUnsignedValue,
    Minimum := FUnsignedMinimum,
    Maximum := FUnsignedMaximum);
END_METHOD

{region 'Documentation'}
(*!
<summary>Checks one subject finding in call order; expected outcomes come from the scenario.</summary>
*)
{endregion}
METHOD PRIVATE CheckFinding : BOOL //! TRUE when the required finding checks pass; calls requiring no finding also succeed.
VAR_INPUT
    Subject : I_Assertion; //! Assertion interface supplying the expected finding identity.
    ExpectedResult : E_Result; //! Independently authored result expected in the captured finding.
    ExpectedFinding : BOOL; //! TRUE when this scenario requires a finding during active evaluation.
END_VAR
VAR_IN_OUT
    Index : UINT; //! One-based next finding index; advanced when this call checks a required finding.
END_VAR
CheckFinding := TRUE;
IF FEvaluateSubjects AND ExpectedFinding THEN
    CheckFinding := (FEvents[Index].SequenceId = UINT_TO_UDINT(Index))
        AND (FEvents[Index].Name = Subject.Name)
        AND (FEvents[Index].OwnerScope = E_OwnerScope.Assertion)
        AND (FEvents[Index].EventType = E_EventType.Result)
        AND (FEvents[Index].State = E_State.Running)
        AND (FEvents[Index].Result = ExpectedResult)
        AND (FEvents[Index].Message <> '');
    Index := Index + 1;
END_IF;
END_METHOD

{region 'Documentation'}
(*!
<summary>Checks exact finding count and identities; at most one finding per subject.</summary>
*)
{endregion}
METHOD PRIVATE CheckFindings
VAR
    Index : UINT;
    Matches : BOOL;
END_VAR
Index := 1;
FFindingsMatch := TRUE;
Matches := CheckFinding(Subject := FSigned,
    ExpectedResult := FSignedExpectedResult,
    ExpectedFinding := FSignedExpectedFinding,
    Index := Index);
FFindingsMatch := FFindingsMatch AND Matches;
Matches := CheckFinding(Subject := FUnsigned,
    ExpectedResult := FUnsignedExpectedResult,
    ExpectedFinding := FUnsignedExpectedFinding,
    Index := Index);
FFindingsMatch := FFindingsMatch AND Matches;
FFindingsMatch := FFindingsMatch
    AND (FCaptureStatus.SequenceId = UINT_TO_UDINT(Index - 1))
    AND (FCaptureStatus.LostEventCount = 0);
IF FEvaluateSubjects AND (FScenario = ScenarioOutsideRange) THEN
    // SA0175: Fixed byte-substring checks of bounded diagnostic messages; no character offsets.
    {analysis -175}
    FFindingsMatch := FFindingsMatch
        AND (FIND(FEvents[1].Message, 'Minimum = -127') > 0)
        AND (FIND(FEvents[1].Message, 'Actual = -128') > 0)
        AND (FIND(FEvents[2].Message, 'Minimum = 128') > 0)
        AND (FIND(FEvents[2].Message, 'Maximum = 255') > 0)
        AND (FIND(FEvents[2].Message, 'Actual = 127') > 0);
    {analysis +175}
END_IF;
IF FEvaluateSubjects AND (FScenario = ScenarioAboveMaximum) THEN
    // SA0175: Fixed byte-substring checks of bounded diagnostic messages; no character offsets.
    {analysis -175}
    FFindingsMatch := FFindingsMatch
        AND (FIND(FEvents[1].Message, 'Maximum = 254') > 0)
        AND (FIND(FEvents[1].Message, 'Actual = 255') > 0);
    {analysis +175}
END_IF;
END_METHOD

{region 'Documentation'}
(*!
<summary>Rejects incomplete subject, capture or outer Assertion setup.</summary>
*)
{endregion}
METHOD PROTECTED CheckInitialization : BOOL //! TRUE when the inherited initialization check and this concrete fixture check both accept the setup.
CheckInitialization := SUPER^.CheckInitialization();
IF NOT CheckInitialization THEN
    RETURN;
END_IF;

CheckInitialization := FSetupValid
    AND FResults.IsInitialized
    AND FActivity.IsInitialized
    AND FInputs.IsInitialized
    AND FFindings.IsInitialized;
IF NOT CheckInitialization THEN
    EventPublisher.PublishEvent(Event := CreateFrameworkEvent(Name := Name,
        ResourceName := '',
        State := State,
        Severity := E_EventSeverity.Error,
        Message := 'Variant selftest setup failed.'));
END_IF;
END_METHOD

{region 'Documentation'}
(*!
<summary>Verifies input preservation without using the tested comparison algorithm.</summary>
*)
{endregion}
METHOD PRIVATE CheckInputs
FInputsMatch := (FSigned.IN = FSignedValue)
    AND (FSigned.Minimum = FSignedMinimum)
    AND (FUnsigned.IN = FUnsignedValue)
    AND (FUnsigned.Minimum = FUnsignedMinimum)
    AND (FUnsigned.Maximum = FUnsignedMaximum);
END_METHOD

{region 'Documentation'}
(*!
<summary>Checks literal evaluation results, or NotEvaluated on the reset call.</summary>
*)
{endregion}
METHOD PRIVATE CheckResults
IF FEvaluateSubjects THEN
    FResultsMatch := (FSigned.Result = FSignedExpectedResult)
        AND (FUnsigned.Result = FUnsignedExpectedResult);
ELSE
    FResultsMatch := (FSigned.Result = E_Result.NotEvaluated)
        AND (FUnsigned.Result = E_Result.NotEvaluated);
END_IF;
FActivityMatch := (FSigned.Enabled = FSubjectEnable)
    AND (FSigned.ObservationActive = (FEvaluateSubjects AND FSubjectEnable))
    AND (FSigned.EvaluationActive = (FEvaluateSubjects AND FSubjectEnable))
    AND (FUnsigned.Enabled = FSubjectEnable)
    AND (FUnsigned.ObservationActive = (FEvaluateSubjects AND FSubjectEnable))
    AND (FUnsigned.EvaluationActive = (FEvaluateSubjects AND FSubjectEnable));
END_METHOD

{region 'Documentation'}
(*!
<summary>Initializes outer checks and isolates intentional subject findings.</summary>
*)
{endregion}
METHOD PROTECTED Configure
VAR
    Initialized : BOOL;
END_VAR
FPreparationStateCount := 0;
FTestStateCount := 1;
FResults.Initialize(Parent := THIS^,
    AssertionName := 'Results');
FActivity.Initialize(Parent := THIS^,
    AssertionName := 'Activity');
FInputs.Initialize(Parent := THIS^,
    AssertionName := 'Inputs');
FFindings.Initialize(Parent := THIS^,
    AssertionName := 'Findings');
FSetupValid := FCapture.Initialize(Buffer := FEvents,
    FifoControl := FCaptureFifo,
    Status := FCaptureStatus);
FSigned.BindPublisher(Publisher := FCapture);
Initialized := FSigned.Initialize(Parent := THIS^,
    AssertionName := 'Signed');
FSetupValid := FSetupValid AND Initialized;
FUnsigned.BindPublisher(Publisher := FCapture);
Initialized := FUnsigned.Initialize(Parent := THIS^,
    AssertionName := 'Unsigned');
FSetupValid := FSetupValid AND Initialized;
END_METHOD

{region 'Documentation'}
(*!
<summary>Completes abort; no asynchronous resource is owned.</summary>
*)
{endregion}
METHOD PROTECTED ProcessAbort
VAR_INPUT
    Enable : BOOL; //! Phase permission supplied by the owning Test Case; FALSE does not authorize progression, while observation may continue.
END_VAR
IF Enable THEN
    CompleteAbort();
END_IF;
END_METHOD

{region 'Documentation'}
(*!
<summary>Latches this call's checks before progression is permitted.</summary>
*)
{endregion}
METHOD PROTECTED ProcessAssertions
VAR_INPUT
    Enable : BOOL; //! Phase permission supplied by the owning Test Case; FALSE does not authorize progression, while observation may continue.
END_VAR
VAR
    Check : BOOL;
END_VAR
Check := Enable AND FObservationReady;
FResults(Enable := Check,
    State := State,
    IN := FResultsMatch);
FActivity(Enable := Check,
    State := State,
    IN := FActivityMatch);
FInputs(Enable := Check,
    State := State,
    IN := FInputsMatch);
FFindings(Enable := Check,
    State := State,
    IN := FFindingsMatch);
IF Check THEN
    FChecked := TRUE;
END_IF;
END_METHOD

{region 'Documentation'}
(*!
<summary>No Preparation phase is needed.</summary>
*)
{endregion}
METHOD PROTECTED ProcessPreparations
VAR_INPUT
    // SA0033: Required hook; this test has no Preparation phase.
    {attribute 'analysis' := '-33'}
    Enable : BOOL; //! Phase permission supplied by the owning Test Case; FALSE does not authorize progression, while observation may continue.
END_VAR
END_METHOD

